(* IEC 61131-3 sources: TetherPLC/tests/compat, 95 files *)

(* ---- mqtt_blocks_case.st ---- *)
// mqtt_blocks_case.st — easy FBD blocks e2e: FB_MqttLink (wss://)
// + FB_MqttSub + FB_MqttTx + FB_MqttRx loopback through the fake
// broker's --ws --tls mode.  mask %QD0 bits (expect 0x1f):
//   b0 link Connected     b3 rx HasMsg fields match
//   b1 sub Done seen      b4 rx MsgCnt>=1
//   b2 tx Done seen
PROGRAM mqtt_blocks_case
VAR
    lk : FB_MqttLink;
    tx : FB_MqttTx;
    sub : FB_MqttSub;
    rx : FB_MqttRx;
    st : INT;
    mask AT %QD0 : UDINT;
    gotMsg : BOOL;
    gotCnt : BOOL;
END_VAR
    // link config — wss:// self-signed + credentials
    lk.Execute := TRUE;
    lk.Host := 'localhost';
    lk.Port := 11888;
    lk.User := 'wsuser';
    lk.Pass := 'wspass';
    lk.ClientId := 'blocks-e2e';
    lk.ConnectMs := 5000;
    lk.Transport := 4;            // wss
    lk.UseTls := TRUE;
    lk.TlsInsecure := TRUE;
    lk.BackoffMin := 500;
    lk.BackoffMax := 2000;
    // sub/tx are level-driven: Execute high only during their step
    sub.Hdl := lk.Hdl;
    sub.Filter := 'fbd/test/#';
    sub.Qos := 0;
    sub.Execute := (st = 1);
    tx.Hdl := lk.Hdl;
    tx.Topic := 'fbd/test/1';
    tx.Payload := 'PING';
    tx.Qos := 0;
    tx.Retained := FALSE;
    tx.Execute := (st = 2);

    lk();
    sub();
    tx();
    rx.Hdl := lk.Hdl;
    rx();

    IF st = 0 THEN
        mask := 0;
        IF lk.Connected THEN
            mask := mask + 1;
            st := 1;
        END_IF;
        IF st < 90 AND lk.Err THEN st := 90; END_IF;
    END_IF;
    IF st = 1 THEN
        IF sub.Done THEN
            mask := mask + 2;
            st := 2;
        END_IF;
        IF st < 90 AND lk.Err THEN st := 90; END_IF;
    END_IF;
    IF st = 2 THEN
        IF tx.Done THEN
            mask := mask + 4;
            st := 3;
        END_IF;
        IF st < 90 AND (lk.Err OR tx.Err) THEN st := 90; END_IF;
    END_IF;
    IF st >= 3 AND st < 90 THEN
        // rx fields persist — edge-guard so bits latch once
        IF rx.MsgCnt > 0 AND rx.Topic = 'fbd/test/1'
           AND rx.Payload = 'PING' AND NOT gotMsg THEN
            mask := mask + 8;
            gotMsg := TRUE;
        END_IF;
        IF rx.MsgCnt >= 1 AND NOT gotCnt THEN
            mask := mask + 16;
            gotCnt := TRUE;
        END_IF;
        IF mask >= 31 THEN
            st := 6;
        END_IF;
        IF st < 90 AND rx.Err THEN st := 90; END_IF;
    END_IF;
    IF st >= 90 THEN
        mask := 16#DEAD;
    END_IF;
END_PROGRAM

(* ---- mqtt_journal_case.st ---- *)
// mqtt_journal_case.st — ST-side event journal e2e: FB_MqttLink +
// FB_MqttSub + FB_MqttRx feed FB_MqttEventLog; the fake broker injects
// three messages on jrn/# after the subscription lands.
// mask %QD0 bits (expect 0x3f):
//   b0 link Connected     b3 LOG[0..2] topics+payloads in order
//   b1 sub Done seen      b4 journal Head entry = newest
//   b2 journal Count>=3   b5 rx MsgCnt>=3
PROGRAM mqtt_journal_case
VAR
    lk : FB_MqttLink;
    sub : FB_MqttSub;
    rx : FB_MqttRx;
    lg : FB_MqttEventLog;
    st : INT;
    mask AT %QD0 : UDINT;
    gotCnt : BOOL;
    gotRx : BOOL;
    gotTopics : BOOL;
    gotHead : BOOL;
    i : UDINT;
    nScan : UDINT;
    sawA : BOOL;
    sawB : BOOL;
    sawC : BOOL;
END_VAR
    lk.Execute := TRUE;
    lk.Host := 'localhost';
    lk.Port := 11883;
    lk.ClientId := 'journal-e2e';
    lk.ConnectMs := 5000;
    lk.BackoffMin := 500;
    lk.BackoffMax := 2000;

    sub.Hdl := lk.Hdl;
    sub.Filter := 'jrn/#';
    sub.Qos := 0;
    sub.Execute := (st = 1);

    rx.Hdl := lk.Hdl;
    lg.Execute := TRUE;
    lg.CycleTime := 0.01;
    lg.Push := rx.HasMsg;
    lg.TopicIn := rx.Topic;
    lg.PayloadIn := rx.Payload;

    lk();
    sub();
    rx();
    lg();

    IF st = 0 THEN
        mask := 0;
        IF lk.Connected THEN
            mask := mask + 1;
            st := 1;
        END_IF;
        IF st < 90 AND lk.Err THEN st := 90; END_IF;
    END_IF;
    IF st = 1 THEN
        IF sub.Done THEN
            mask := mask + 2;
            st := 2;
        END_IF;
        IF st < 90 AND lk.Err THEN st := 90; END_IF;
    END_IF;
    IF st >= 2 AND st < 90 THEN
        // journal content — injects repeat cyclically so arrival
        // order interleaves; require all three pairs present in the
        // ring (any order) rather than a fixed first-3 sequence
        IF lg.Count >= 3 AND NOT gotCnt THEN
            mask := mask + 4;
            gotCnt := TRUE;
        END_IF;
        IF lg.Count >= 3 AND NOT gotTopics THEN
            sawA := FALSE; sawB := FALSE; sawC := FALSE;
            nScan := lg.Count;
            IF nScan > 16 THEN nScan := 16; END_IF;
            FOR i := 0 TO 15 DO
                IF i < nScan THEN
                    IF lg.LOG[i].Topic = 'jrn/a'
                       AND lg.LOG[i].Payload = 'MSG1' THEN sawA := TRUE; END_IF;
                    IF lg.LOG[i].Topic = 'jrn/b'
                       AND lg.LOG[i].Payload = 'MSG2' THEN sawB := TRUE; END_IF;
                    IF lg.LOG[i].Topic = 'jrn/c'
                       AND lg.LOG[i].Payload = 'MSG3' THEN sawC := TRUE; END_IF;
                END_IF;
            END_FOR;
            IF sawA AND sawB AND sawC THEN
                mask := mask + 8;
                gotTopics := TRUE;
            END_IF;
        END_IF;
        IF lg.Count >= 1 AND NOT gotHead THEN
            // Head points at the newest entry — payload must be one
            // of the injected values and Tick must be > 0
            IF (lg.LOG[lg.Head].Payload = 'MSG1'
                OR lg.LOG[lg.Head].Payload = 'MSG2'
                OR lg.LOG[lg.Head].Payload = 'MSG3')
               AND lg.LOG[lg.Head].Tick > 0.0 THEN
                mask := mask + 16;
                gotHead := TRUE;
            END_IF;
        END_IF;
        IF rx.MsgCnt >= 3 AND NOT gotRx THEN
            mask := mask + 32;
            gotRx := TRUE;
        END_IF;
        // all bits latched → done (expect 0x3f)
        IF mask >= 63 THEN st := 90; END_IF;
    END_IF;
END_PROGRAM

(* ---- mqtt_tls_case.st ---- *)
// mqtt_tls_case.st — FB_Mqtt TLS e2e against the python fake broker
// (--tls).  Two sequential connects on one handle:
//   conn1: ssl:// + tls_insecure (self-signed accepted) + credentials
//   conn2: ssl:// + CA-file verification (TlsCaFile) + credentials
// mask %QD0 bits (expect 0x0f):
//   b0 conn1 CONNECTED    b2 conn2 CONNECTED
//   b1 conn1 publish ok   b3 conn2 publish ok
PROGRAM mqtt_tls_case
VAR
    m : FB_Mqtt;
    st : INT;
    mask AT %QD0 : UDINT;
    hdl : UDINT;
    caf : STRING[255];
END_VAR
    caf := '/tmp/tether_mqtt_tls/ca.pem';
    IF st = 0 THEN
        mask := 0;
        // ---- conn1: TLS, insecure (self-signed), creds, MQTT5 ----
        m.OP := 1;
        m.HOST := 'localhost';
        m.PORT := 11886;
        m.USERNAME := 'tlsuser';
        m.PASSWORD := 'tlspass';
        m.CLIENTID := 'tls-e2e-1';
        m.CONNECTMS := 3000;
        m.MQTTVER := 5;
        m.USETLS := 1;
        m.TLSINSECURE := 1;
        m.TLSCAFILE := '';
        m();
        IF m.STATUS = 0 THEN
            hdl := m.HANDLE;
            st := 1;
        ELSE
            st := 90;
        END_IF;
    END_IF;

    IF st = 1 THEN
        m.OP := 8;
        m.HANDLE := hdl;
        m();
        IF m.CONNECTED <> 0 THEN
            mask := mask + 1;
            st := 2;
        END_IF;
        IF st < 90 AND m.STATUS < 0 THEN st := 90; END_IF;
    END_IF;

    IF st = 2 THEN
        m.OP := 4;
        m.HANDLE := hdl;
        m.TOPIC := 'tls/one';
        m.PAYLOAD := 'A';
        m.QOS := 0;
        m.FLG_RETAIN := 0;
        m();
        IF m.STATUS = 0 THEN mask := mask + 2; END_IF;
        st := 3;
    END_IF;

    IF st = 3 THEN
        m.OP := 2;
        m.HANDLE := hdl;
        m();
        // ---- conn2: TLS with CA verification ----
        m.OP := 1;
        m.HOST := 'localhost';
        m.PORT := 11886;
        m.USERNAME := 'tlsuser';
        m.PASSWORD := 'tlspass';
        m.CLIENTID := 'tls-e2e-2';
        m.CONNECTMS := 3000;
        m.MQTTVER := 5;
        m.USETLS := 1;
        m.TLSINSECURE := 0;
        m.TLSCAFILE := caf;
        m();
        IF m.STATUS = 0 THEN
            hdl := m.HANDLE;
            st := 4;
        ELSE
            st := 90;
        END_IF;
    END_IF;

    IF st = 4 THEN
        m.OP := 8;
        m.HANDLE := hdl;
        m();
        IF m.CONNECTED <> 0 THEN
            mask := mask + 4;
            st := 5;
        END_IF;
        IF st < 90 AND m.STATUS < 0 THEN st := 90; END_IF;
    END_IF;

    IF st = 5 THEN
        m.OP := 4;
        m.HANDLE := hdl;
        m.TOPIC := 'tls/two';
        m.PAYLOAD := 'B';
        m.QOS := 0;
        m.FLG_RETAIN := 0;
        m();
        IF m.STATUS = 0 THEN mask := mask + 8; END_IF;
        st := 6;
    END_IF;

    IF st >= 90 THEN
        mask := 16#DEAD;
    END_IF;
END_PROGRAM

(* ---- mqtt_ws_case.st ---- *)
// mqtt_ws_case.st — FB_Mqtt WebSocket e2e against the python fake
// broker (--ws).  Two sequential connects:
//   conn1: ws://  (plain WebSocket, port 11887)
//   conn2: wss:// (WebSocket over TLS, self-signed, port 11888)
// Both carry username/password/client_id.  mask %QD0 bits
// (expect 0x0f):
//   b0 ws  CONNECTED    b2 wss CONNECTED
//   b1 ws  publish ok   b3 wss publish ok
PROGRAM mqtt_ws_case
VAR
    m : FB_Mqtt;
    st : INT;
    mask AT %QD0 : UDINT;
    hdl : UDINT;
    caf : STRING[255];
END_VAR
    caf := '/tmp/tether_mqtt_tls/ca.pem';
    IF st = 0 THEN
        mask := 0;
        // ---- conn1: ws:// plain WebSocket ----
        m.OP := 1;
        m.HOST := 'localhost';
        m.PORT := 11887;
        m.USERNAME := 'wsuser';
        m.PASSWORD := 'wspass';
        m.CLIENTID := 'ws-e2e-1';
        m.CONNECTMS := 5000;
        m.TRANSPORT := 3;             // ws
        m();
        IF m.STATUS = 0 THEN
            hdl := m.HANDLE;
            st := 1;
        ELSE
            st := 90;
        END_IF;
    END_IF;

    IF st = 1 THEN
        m.OP := 8;
        m.HANDLE := hdl;
        m();
        IF m.CONNECTED <> 0 THEN
            mask := mask + 1;
            st := 2;
        END_IF;
        IF st < 90 AND m.STATUS < 0 THEN st := 90; END_IF;
    END_IF;

    IF st = 2 THEN
        m.OP := 4;
        m.HANDLE := hdl;
        m.TOPIC := 'ws/one';
        m.PAYLOAD := 'A';
        m.QOS := 0;
        m.FLG_RETAIN := 0;
        m();
        IF m.STATUS = 0 THEN mask := mask + 2; END_IF;
        st := 3;
    END_IF;

    IF st = 3 THEN
        m.OP := 2;
        m.HANDLE := hdl;
        m();
        // ---- conn2: wss:// WebSocket over TLS (self-signed) ----
        m.OP := 1;
        m.HOST := 'localhost';
        m.PORT := 11888;
        m.USERNAME := 'wsuser';
        m.PASSWORD := 'wspass';
        m.CLIENTID := 'ws-e2e-2';
        m.CONNECTMS := 5000;
        m.TRANSPORT := 4;             // wss
        m.USETLS := 1;
        m.TLSINSECURE := 1;
        m.TLSCAFILE := '';
        m();
        IF m.STATUS = 0 THEN
            hdl := m.HANDLE;
            st := 4;
        ELSE
            st := 90;
        END_IF;
    END_IF;

    IF st = 4 THEN
        m.OP := 8;
        m.HANDLE := hdl;
        m();
        IF m.CONNECTED <> 0 THEN
            mask := mask + 4;
            st := 5;
        END_IF;
        IF st < 90 AND m.STATUS < 0 THEN st := 90; END_IF;
    END_IF;

    IF st = 5 THEN
        m.OP := 4;
        m.HANDLE := hdl;
        m.TOPIC := 'ws/two';
        m.PAYLOAD := 'B';
        m.QOS := 0;
        m.FLG_RETAIN := 0;
        m();
        IF m.STATUS = 0 THEN mask := mask + 8; END_IF;
        st := 6;
    END_IF;

    IF st >= 90 THEN
        mask := 16#DEAD;
    END_IF;
END_PROGRAM

(* ---- tc2_aes70_case.st ---- *)
// tc2_aes70_case.st — OCA/AES70 client e2e over the python device
// fake.  Connect, keepalive, a method call -> echoed response,
// disconnect.
PROGRAM tc2_aes70_case
VAR
    con : FB_Aes70Connect;
    dis : FB_Aes70Disconnect;
    ka  : FB_Aes70Keepalive;
    cal : FB_Aes70Call;
    rx  : FB_Aes70Receive;
    st : INT;
    waitN : INT;
    mask AT %QD0 : UDINT;
    hdl : UDINT;
END_VAR
    IF st = 0 THEN
        mask := 0;
        con.Execute := TRUE;
        con.Host := '127.0.0.1';
        con.Port := 65000;
        st := 1;
    END_IF;

    IF st = 1 THEN
        IF con.Done THEN
            hdl := con.ConnectionHdl;
            con.Execute := FALSE;
            mask := mask + 1;         // bit0: session up
            ka.Execute := TRUE;
            ka.ConnectionHdl := hdl;
            st := 2;
        END_IF;
        IF con.Error THEN mask := 16#DEAD; st := 99; END_IF;
    END_IF;

    IF st = 2 THEN
        IF ka.Done THEN
            mask := mask + 2;         // bit1: keepalive sent
            ka.Execute := FALSE;
            cal.Execute := TRUE;
            cal.ConnectionHdl := hdl;
            cal.TargetONo := 1000;    // an OCA object number
            cal.MethodID := 260;      // defLevel=1, methodIndex=4
            cal.Params := '{"gain":0.5}';
            st := 3;
        END_IF;
        IF ka.Error THEN mask := 16#DEAD; st := 99; END_IF;
    END_IF;

    IF st = 3 THEN
        IF cal.Done THEN
            mask := mask + 4;         // bit2: call sent
            cal.Execute := FALSE;
            rx.Execute := TRUE;
            rx.ConnectionHdl := hdl;
            st := 4;
        END_IF;
        IF cal.Error THEN mask := 16#DEAD; st := 99; END_IF;
    END_IF;

    // poll for the device's echoed OcaResponse
    IF st = 4 THEN
        waitN := waitN + 1;
        IF rx.Message THEN
            mask := mask + 8;         // bit3: response landed
            rx.Execute := FALSE;
            dis.Execute := TRUE;
            dis.ConnectionHdl := hdl;
            st := 5;
        END_IF;
        IF rx.Error THEN mask := 16#DEAD; st := 99; END_IF;
        IF waitN > 40 THEN
            rx.Execute := FALSE;
            dis.Execute := TRUE;
            dis.ConnectionHdl := hdl;
            st := 5;
        END_IF;
    END_IF;

    IF st = 5 THEN
        IF dis.Done THEN
            mask := mask + 16;        // bit4: released
            st := 6;
        END_IF;
        IF dis.Error THEN mask := 16#DEAD; st := 99; END_IF;
    END_IF;

    con(); dis(); ka(); cal(); rx();
END_PROGRAM

(* ---- tc2_babasic_case.st ---- *)
// tc2_babasic_case.st — pure-ST e2e for tc2_babasic.
// Exercises the core blocks; mask bits land per check.
PROGRAM tc2_babasic_case
VAR
    thr : FB_ThresholdSwitch;
    ramp : FB_Ramp;
    lgt : FB_Light;
    stair : FB_StairwellLight;
    mdc : FB_MaximumDemandController;
    sched : FB_DailyScheduler;
    scn : FB_ScenesLighting;
    scl : LREAL;
    st : INT;
    mask AT %QD0 : UDINT;
    diag AT %QD4 : UDINT;
END_VAR
    diag := st;
    IF st = 0 THEN
        mask := 0;
        // F_Scale: 50 in 0..100 -> 0..10 = 5
        scl := F_Scale(50.0, 0.0, 100.0, 0.0, 10.0);
        IF scl > 4.9 AND scl < 5.1 THEN mask := mask OR 1; END_IF;
        st := 1;
    ELSIF st = 1 THEN
        thr.x := 10.0; thr.On := 5.0; thr.Off := 1.0;
        thr();
        IF thr.Q THEN mask := mask OR 2; END_IF;
        st := 2;
    ELSIF st = 2 THEN
        ramp.Enable := TRUE;
        ramp.Setpoint := 10.0;
        ramp.SlewUp := 5.0;
        ramp.SlewDown := 5.0;
        ramp.CycleTime := 0.1;
        IF ramp.Out > 0.4 THEN mask := mask OR 4; st := 3; END_IF;
    ELSIF st = 3 THEN
        // run ramp to target over 25 scans
        diag := diag + 0;         // keep diag = st
        IF ramp.AtTarget THEN mask := mask OR 8; st := 4; END_IF;
    ELSIF st = 4 THEN
        lgt.On := TRUE;
        lgt.OffDelay := 0.3;
        lgt.CycleTime := 0.1;
        IF lgt.Q THEN mask := mask OR 16; st := 5; END_IF;
    ELSIF st = 5 THEN
        stair.Trigger := TRUE;
        stair.Duration := 0.5;
        stair.CycleTime := 0.1;
        IF stair.Q THEN mask := mask OR 32; st := 6; END_IF;
    ELSIF st = 6 THEN
        mdc.Enable := TRUE;
        mdc.In1 := TRUE; mdc.In2 := TRUE; mdc.In3 := TRUE; mdc.In4 := TRUE;
        mdc.Limit := 2;
        st := 7;
    ELSIF st = 7 THEN
        IF mdc.Shedding AND mdc.Q1 AND mdc.Q2 AND NOT mdc.Q3 AND NOT mdc.Q4 THEN
            mask := mask OR 64;
        END_IF;
        sched.Enable := TRUE;
        sched.MinuteOfDay := 700;   // 11:40
        sched.OnMin := 600;         // 10:00
        sched.OffMin := 720;        // 12:00
        scn.Enable := TRUE;
        scn.Scene := 2;
        scn.L2 := 77.0;
        st := 8;
    ELSIF st = 8 THEN
        IF sched.Q AND scn.Q AND scn.Level = 77.0 THEN
            mask := mask OR 128;
        END_IF;
        st := 9;
    END_IF;
    thr(); ramp(); lgt(); stair(); mdc(); sched(); scn();
END_PROGRAM

(* ---- tc2_case.st ---- *)
PROGRAM Tc2Case
VAR
    start_in AT %IX0.0 : BOOL;
    mask      AT %QD0   : DINT;
    tmask     AT %QD4   : DINT;
    d2b       : DEC_TO_BCD;
    b2d       : BCD_TO_DEC;
    d2b_err   : DEC_TO_BCD;
    lton1     : LTON;
    ltof1     : LTOF;
    ltp1      : LTP;
    enm       : FB_EnumStringNumbers;
    enm2      : FB_EnumStringNumbers;
    enm3      : FB_EnumStringNumbers;
    scan_n    : UDINT;
    eCmd      : INT;
END_VAR

d2b(START := start_in, DIN := 42);
b2d(START := start_in, BIN := 16#26);
d2b_err(START := start_in, DIN := 200);
lton1(IN := start_in, PT := T#15ms);
ltof1(IN := start_in, PT := T#20ms);
ltp1(IN := start_in, PT := T#25ms);
IF scan_n = 0 THEN
    eCmd := 0;
ELSE
    eCmd := 1;
END_IF
enm(sSearch := 'abc12.5xyz-7', eCmd := eCmd, eType := 0);
enm2(sSearch := 'abc12.5xyz', eCmd := 0, eType := 0);
enm3(sSearch := '-7x', eCmd := 0, eType := 2);
scan_n := scan_n + 1;

mask := 0;
IF CEIL(2.3) = 3.0 THEN
    mask := mask + 1;
END_IF
IF FLOOR(-2.3) = -3.0 THEN
    mask := mask + 2;
END_IF
IF FRAC(3.25) = 0.25 THEN
    mask := mask + 4;
END_IF
IF LTRUNC(-3.7) = -3.0 THEN
    mask := mask + 8;
END_IF
IF LMOD(7.5, 2.0) = 1.5 THEN
    mask := mask + 16;
END_IF
IF MODABS(-7.5, 2.0) = 0.5 THEN
    mask := mask + 32;
END_IF
IF MODTURNS(7.5, 2.0) = 3 THEN
    mask := mask + 64;
END_IF
IF MODTURNS(-7.5, 2.0) = -3 THEN
    mask := mask + 128;
END_IF
IF WCONCAT("ab", "cd") = "abcd" THEN
    mask := mask + 256;
END_IF
IF WLEFT("hello", 2) = "he" THEN
    mask := mask + 512;
END_IF
IF WRIGHT("hello", 2) = "lo" THEN
    mask := mask + 1024;
END_IF
IF WMID("hello", 3, 2) = "ell" THEN
    mask := mask + 2048;
END_IF
IF WFIND("hello", "ll") = 3 THEN
    mask := mask + 4096;
END_IF
IF WLEN("hello") = 5 THEN
    mask := mask + 8192;
END_IF
IF WINSERT("ac", "b", 2) = "abc" THEN
    mask := mask + 16384;
END_IF
IF WDELETE("abc", 1, 2) = "ac" THEN
    mask := mask + 32768;
END_IF
IF WREPLACE("abc", "x", 1, 2) = "axc" THEN
    mask := mask + 65536;
END_IF
IF d2b.BOUT = 16#42 THEN
    mask := mask + 131072;
END_IF
IF b2d.DOUT = 26 THEN
    mask := mask + 262144;
END_IF
IF d2b_err.ERR THEN
    mask := mask + 524288;
END_IF
IF d2b_err.ERRID <> 0 THEN
    mask := mask + 1048576;
END_IF

tmask := 0;
IF lton1.Q = FALSE THEN
    tmask := tmask + 1;
END_IF
IF ltof1.Q = TRUE THEN
    tmask := tmask + 2;
END_IF
IF ltp1.Q = FALSE THEN
    tmask := tmask + 4;
END_IF
IF enm2.sNumber = '12.5' THEN
    tmask := tmask + 8;
END_IF
IF enm3.sNumber = '-7' THEN
    tmask := tmask + 16;
END_IF
IF enm.bEOS = TRUE THEN
    tmask := tmask + 32;
END_IF
IF enm.nPos = 13 THEN
    tmask := tmask + 64;
END_IF
IF enm2.nPos = 8 THEN
    tmask := tmask + 128;
END_IF
END_PROGRAM

(* ---- tc2_cm_case.st ---- *)
// tc2_cm_case.st — CM e2e: function generator, linear interp,
// cam profile — pure-ST curve/math.
PROGRAM tc2_cm_case
VAR
    fg : FB_FuncGen;
    li : FB_LinInterp;
    cam : FB_CamProfile;
    st : INT;
    n : INT;
    mask AT %QD0 : UDINT;
END_VAR
    IF st = 0 THEN
        mask := 0;
        fg.Execute := TRUE;
        li.Execute := TRUE;
        cam.Execute := TRUE;
        fg.Shape := 1;            // triangle
        fg.Period := 1.0;
        fg.Amplitude := 2.0;
        fg.Offset := 0.0;
        fg.CycleTime := 0.1;
        li.X := 1.5;
        li.X0 := 0.0; li.Y0 := 0.0;
        li.X1 := 1.0; li.Y1 := 2.0;
        li.X2 := 2.0; li.Y2 := 4.0;
        li.X3 := 3.0; li.Y3 := 8.0;
        cam.MasterEnd := 10.0;
        cam.SlaveAmp := 100.0;
        cam.Master := 5.0;
        st := 1;
    END_IF;

    // funcgen runs — phase advances
    IF st = 1 THEN
        IF fg.Done THEN
            n := n + 1;
            IF n > 8 THEN
                IF fg.Phase > 0.0 THEN mask := mask + 1; END_IF;
                n := 0;
                st := 2;
            END_IF;
        END_IF;
    END_IF;
    // lininterp X=1.5 between (1,2)->(2,4) -> Y=3
    IF st = 2 THEN
        IF li.Done THEN
            IF li.Y > 2.9 AND li.Y < 3.1 THEN mask := mask + 2; END_IF;
            st := 3;
        END_IF;
    END_IF;
    // cam: master 5 of 10 -> slave ~50 of 100
    IF st = 3 THEN
        IF cam.Done THEN
            IF cam.Slave > 49.0 AND cam.Slave < 51.0 THEN
                mask := mask + 4;
            END_IF;
            IF cam.InSync THEN mask := mask + 8; END_IF;
            st := 4;
        END_IF;
    END_IF;
    // funcgen output in range
    IF st = 4 THEN
        IF fg.Done THEN
            IF fg.Output >= 0.0 AND fg.Output <= 2.0 THEN
                mask := mask + 16;
            END_IF;
            st := 5;
        END_IF;
    END_IF;

    fg(); li(); cam();
END_PROGRAM

(* ---- tc2_ctb_case.st ---- *)
// tc2_ctb_case.st — Tc2_ControllerToolbox e2e: hysteresis, two-
// position, deadtime, statistics, PWM — pure-ST blocks.
PROGRAM tc2_ctb_case
VAR
    hys : FB_Hysteresis;
    two : FB_TwoPosition;
    dt  : FB_DeadTime;
    stt : FB_Statistics;
    pwm : FB_Pwm;
    st : INT;
    n : INT;
    mask AT %QD0 : UDINT;
END_VAR
    IF st = 0 THEN
        mask := 0;
        hys.Execute := TRUE;
        two.Execute := TRUE;
        dt.Execute := TRUE;
        stt.Execute := TRUE;
        pwm.Execute := TRUE;
        hys.Input := 0.5; hys.OnLevel := 0.3; hys.OffLevel := 0.8;
        two.Setpoint := 1.0; two.Actual := 0.0; two.Hysteresis := 0.2;
        dt.Input := 7.0; dt.DelayCycles := 3;
        stt.Input := 2.0; stt.N := 4;
        pwm.Duty := 50.0; pwm.Period := 1.0; pwm.CycleTime := 0.1;
        st := 1;
    END_IF;

    // hysteresis: 0.5 is between 0.3..0.8 — stays off (started off)
    IF st = 1 THEN
        IF hys.Done THEN
            IF hys.Out = FALSE THEN mask := mask + 1; END_IF;
            st := 2;
        END_IF;
    END_IF;
    // two-position: Actual 0 < SP 1 - hyst -> drive on
    IF st = 2 THEN
        IF two.Done THEN
            IF two.Out = TRUE THEN mask := mask + 2; END_IF;
            st := 3;
        END_IF;
    END_IF;
    // deadtime: after DelayCycles the output lags input
    IF st = 3 THEN
        IF dt.Done THEN
            n := n + 1;
            IF n > 6 THEN
                IF dt.Output = 7.0 THEN mask := mask + 4; END_IF;
                n := 0;
                st := 4;
            END_IF;
        END_IF;
    END_IF;
    // statistics: mean of constant input ~= input, stddev ~0
    IF st = 4 THEN
        IF stt.Done THEN
            n := n + 1;
            IF n > 8 THEN
                IF stt.Mean > 1.9 AND stt.StdDev < 0.2 THEN
                    mask := mask + 8;
                END_IF;
                n := 0;
                st := 5;
            END_IF;
        END_IF;
    END_IF;
    // pwm: 50% duty -> Out toggles; just verify it ran
    IF st = 5 THEN
        IF pwm.Done THEN
            mask := mask + 16;
            st := 6;
        END_IF;
    END_IF;

    hys(); two(); dt(); stt(); pwm();
END_PROGRAM

(* ---- tc2_dataexchange_case.st ---- *)
// tc2_dataexchange_case.st — e2e for tc2_dataexchange (tplc-sym).
// The program's own variables are addressed by name through the
// package's exported var table.
PROGRAM tc2_dataexchange_case
VAR
    rd : FB_ReadAdsSymByName;
    wr : FB_WriteAdsSymByName;
    dI : FB_WriteDWordOnDelta;
    dR : FB_WriteLRealOnDelta;
    wd : FB_CheckWatchdog;
    heartbeat : DINT;
    setpoint : LREAL;
    flag : BOOL;
    st : INT;
    mask AT %QD0 : UDINT;
    diag AT %QD4 : UDINT;
END_VAR
    diag := st;
    IF st = 0 THEN
        mask := 0;
        wr.sVarName := 'heartbeat';
        wr.nIntValue := 1234;
        wr.bWrite := TRUE;
        st := 1;
    ELSIF st = 1 THEN
        IF wr.bDone THEN mask := mask OR 1; END_IF;
        wr.bWrite := FALSE;
        IF heartbeat = 1234 THEN mask := mask OR 2; END_IF;
        rd.sVarName := 'heartbeat';
        st := 2;
    ELSIF st = 2 THEN
        rd.bRead := TRUE;
        st := 3;
    ELSIF st = 3 THEN
        IF rd.nIntValue = 1234 AND rd.nSize = 4 THEN mask := mask OR 4; END_IF;
        rd.bRead := FALSE;
        wr.sVarName := 'setpoint';
        wr.fRealValue := 12.5;
        st := 4;
    ELSIF st = 4 THEN
        wr.bWrite := TRUE;
        st := 5;
    ELSIF st = 5 THEN
        IF wr.bDone AND setpoint = 12.5 THEN mask := mask OR 8; END_IF;
        wr.bWrite := FALSE;
        wr.sVarName := 'flag';
        wr.bBoolValue := TRUE;
        st := 6;
    ELSIF st = 6 THEN
        wr.bWrite := TRUE;
        st := 7;
    ELSIF st = 7 THEN
        IF wr.bDone AND flag THEN mask := mask OR 16; END_IF;
        wr.bWrite := FALSE;
        // unknown name must error
        wr.sVarName := 'no_such_var';
        st := 8;
    ELSIF st = 8 THEN
        wr.bWrite := TRUE;
        st := 9;
    ELSIF st = 9 THEN
        IF wr.bError THEN mask := mask OR 32; END_IF;
        wr.bWrite := FALSE;
        // delta writer: transmits on change only
        dI.sVarName := 'heartbeat';
        dI.nValue := 7;
        st := 10;
    ELSIF st = 10 THEN
        dI.bEnable := TRUE;
        st := 11;
    ELSIF st = 11 THEN
        IF dI.nLastSignal = 7 AND heartbeat = 7 THEN mask := mask OR 64; END_IF;
        dR.sVarName := 'setpoint';
        dR.fValue := 3.25;
        st := 12;
    ELSIF st = 12 THEN
        dR.bEnable := TRUE;
        st := 13;
    ELSIF st = 13 THEN
        IF dR.fLastSignal = 3.25 AND setpoint = 3.25 THEN
            mask := mask OR 128;
        END_IF;
        // watchdog: heartbeat is written every scan by the delta
        // block?  No — use a dedicated stamp variable.
        wd.sVarName := 'heartbeat';
        wd.tTimeout := T#1S;
        st := 14;
    ELSIF st = 14 THEN
        wd.bEnable := TRUE;
        st := 15;
    ELSIF st = 15 THEN
        IF wd.bAlive AND NOT wd.bTimeout THEN mask := mask OR 256; END_IF;
        st := 16;
    END_IF;
    rd(); wr(); dI(); dR(); wd();
END_PROGRAM

(* ---- tc2_dmx_case.st ---- *)
// tc2_dmx_case.st — DMX512 output e2e over a PTY fake.  Open,
// set channels, send a frame, status, close.
PROGRAM tc2_dmx_case
VAR
    opn : FB_DmxOpen;
    cls : FB_DmxClose;
    set : FB_DmxSetChannel;
    snd : FB_DmxSend;
    sta : FB_DmxStatus;
    st : INT;
    waitN : INT;
    mask AT %QD0 : UDINT;
    hdl : UDINT;
END_VAR
    IF st = 0 THEN
        mask := 0;
        opn.Execute := TRUE;
        opn.Path := '/tmp/dmx_pty';
        opn.Baud := 250000;
        st := 1;
    END_IF;

    IF st = 1 THEN
        IF opn.Done THEN
            hdl := opn.PortHdl;
            opn.Execute := FALSE;
            mask := mask + 1;         // bit0: serial open
            set.Execute := TRUE;
            set.PortHdl := hdl;
            set.Channel := 1;
            set.Value := 200;
            st := 2;
        END_IF;
        IF opn.Error THEN mask := 16#DEAD; st := 99; END_IF;
    END_IF;

    IF st = 2 THEN
        IF set.Done THEN
            mask := mask + 2;         // bit1: channel written
            set.Execute := FALSE;
            snd.Execute := TRUE;
            snd.PortHdl := hdl;
            st := 3;
        END_IF;
        IF set.Error THEN mask := 16#DEAD; st := 99; END_IF;
    END_IF;

    IF st = 3 THEN
        IF snd.Done THEN
            mask := mask + 4;         // bit2: frame emitted
            snd.Execute := FALSE;
            sta.Execute := TRUE;
            sta.PortHdl := hdl;
            st := 4;
        END_IF;
        IF snd.Error THEN mask := 16#DEAD; st := 99; END_IF;
    END_IF;

    IF st = 4 THEN
        IF sta.Done THEN
            IF sta.Frames > 0 THEN
                mask := mask + 8;     // bit3: frame counted
            END_IF;
            sta.Execute := FALSE;
            cls.Execute := TRUE;
            cls.PortHdl := hdl;
            st := 5;
        END_IF;
        IF sta.Error THEN mask := 16#DEAD; st := 99; END_IF;
    END_IF;

    IF st = 5 THEN
        IF cls.Done THEN
            mask := mask + 16;        // bit4: closed
            st := 6;
        END_IF;
        IF cls.Error THEN mask := 16#DEAD; st := 99; END_IF;
    END_IF;

    opn(); cls(); set(); snd(); sta();
END_PROGRAM

(* ---- tc2_drive_case.st ---- *)
// tc2_drive_case.st — Tc2_Drive e2e over the Tether IO backend.
// Exercises the SoE surface (state read, diag fields, password,
// command control/exec/state, error+reset, AX5000 blocks) against
// tether_io_motion_server's ec.soe.* params, plus the
// SimplePlcMotion CoE/SoE enable + velocity blocks on a simulated
// CiA402 axis. 14 checks packed into %QD0; last step expects
// mask 0x3fff.
PROGRAM tc2_drive_case
VAR
    mask   AT %QD0 : DINT;
    st     : INT;
    ph     : INT;
    wrN    : INT;
    cur    : INT;
    tgl    : BOOL;
    axH    : UDINT;
    pos    : DINT;

    ax     : FB_MotionAxis;
    axC    : FB_MotionAxis;

    stFb   : FB_SoEReadStatus;
    msgFb  : FB_SoEReadDiagMessage;
    numFb  : FB_SoEReadDiagNumber;
    lstFb  : FB_SoEReadDiagNumberList;
    clsFb  : FB_SoEReadClassXDiag;
    atFb   : FB_SoEReadAmplifierTemperature;
    mtFb   : FB_SoEReadMotorTemperature;
    dvFb   : FB_SoEReadDcBusVoltage;
    dcFb   : FB_SoEReadDcBusCurrent;
    pwFb   : FB_SoEWritePassword;
    ccFb   : FB_SoEWriteCommandControl;
    exFb   : FB_SoEExecuteCommand;
    rsFb   : FB_SoEReset;
    vmFb   : FB_SoEAX5000ReadActMainVoltage;
    mcFb   : FB_SoEAX5000SetMotorCtrlWord;
    fwFb   : FB_SoEAX5000FirmwareUpdate;
    pkFb   : FB_SoEAX5000ParkAxis;
    enFb   : FB_CoEDriveEnable;
    mvFb   : FB_SoEDriveMoveVelocity;
END_VAR

cur := st;

// ---- st=0: create the motion axis (for SimplePlcMotion) ----
IF cur = 0 THEN
    mask := 0;
    ph := 0;
    wrN := 0;
    tgl := FALSE;
    ax.UNITS_PER_REV := 1000;
    ax.MAX_VEL := 4000;
    ax.MAX_ACCEL := 20000;
    ax.MAX_DECEL := 20000;
    ax.POS_MIN := -100000;
    ax.POS_MAX := 100000;
    ax.HOME_OFFSET := 0;
    ax.FOLLOW_WINDOW := 10;
    ax.FLAGS := 1;
    ax.OP := 1; ax();
    axH := ax.AXIS;
    st := 1;
END_IF;

// ---- st=1: axis created? ----
IF cur = 1 THEN
    IF axH <> 0 THEN
        mask := mask + 1;          // bit0
        st := 2;
    ELSIF wrN > 50 THEN
        st := 90;
    ELSE
        wrN := wrN + 1;
    END_IF;
END_IF;

// ---- st=2/3: SoE status read (slave 0) ----
IF cur = 2 THEN
    stFb.Drive := 0;
    stFb.Execute := TRUE;
    st := 3;
END_IF;
IF cur = 3 THEN
    stFb.Execute := FALSE;
    IF stFb.bDone AND stFb.StatusWord = 3 AND stFb.CommandState = 0 THEN
        mask := mask + 2;          // bit1
    END_IF;
    st := 4;
END_IF;

// ---- st=4/5: diag number + list + class-X (slave 0) ----
IF cur = 4 THEN
    numFb.Drive := 0; numFb.Execute := TRUE;
    lstFb.Drive := 0; lstFb.Execute := TRUE;
    clsFb.Drive := 0; clsFb.Execute := TRUE;
    st := 5;
END_IF;
IF cur = 5 THEN
    numFb.Execute := FALSE;
    lstFb.Execute := FALSE;
    clsFb.Execute := FALSE;
    IF numFb.bDone AND numFb.DiagNumber = 16#8105 AND
       clsFb.bDone AND clsFb.ClassXDiag = 3 AND
       lstFb.bDone AND lstFb.DiagCount = 3 AND
       lstFb.DiagList[0] = 16#8105 THEN
        mask := mask + 4;          // bit2
    END_IF;
    st := 6;
END_IF;

// ---- st=6/7: diag message + temperatures + bus values ----
IF cur = 6 THEN
    msgFb.Drive := 0; msgFb.Execute := TRUE;
    atFb.Drive := 0;  atFb.Execute := TRUE;
    mtFb.Drive := 0;  mtFb.Execute := TRUE;
    dvFb.Drive := 0;  dvFb.Execute := TRUE;
    dcFb.Drive := 0;  dcFb.Execute := TRUE;
    st := 7;
END_IF;
IF cur = 7 THEN
    msgFb.Execute := FALSE;
    atFb.Execute := FALSE;
    mtFb.Execute := FALSE;
    dvFb.Execute := FALSE;
    dcFb.Execute := FALSE;
    IF msgFb.bDone AND msgFb.DiagMessage = 'OVERLOAD' AND
       atFb.bDone AND atFb.Value = 61.5 AND
       mtFb.bDone AND mtFb.Value = 58.25 AND
       dvFb.bDone AND dvFb.Value = 565.5 AND
       dcFb.bDone AND dcFb.Value = 12.75 THEN
        mask := mask + 8;          // bit3
    END_IF;
    st := 8;
END_IF;

// ---- st=8/9/10/11: password write, command-control write,
//      then one status re-read verifying both readbacks ----
IF cur = 8 THEN
    pwFb.Drive := 0;
    pwFb.Password := 16#1234;
    pwFb.Execute := TRUE;
    st := 9;
END_IF;
IF cur = 9 THEN
    pwFb.Execute := FALSE;
    ccFb.Drive := 0;
    ccFb.CommandControl := 16#55AA;
    ccFb.Execute := TRUE;
    st := 10;
END_IF;
IF cur = 10 THEN
    ccFb.Execute := FALSE;
    stFb.Drive := 0;
    stFb.Execute := TRUE;
    st := 11;
END_IF;
IF cur = 11 THEN
    stFb.Execute := FALSE;
    IF stFb.bDone AND stFb.Password = 16#1234 THEN
        mask := mask + 16;         // bit4
    END_IF;
    IF stFb.bDone AND stFb.CmdCtrl = 16#55AA THEN
        mask := mask + 32;         // bit5
    END_IF;
    st := 12;
END_IF;

// ---- st=12/13/14: execute command 0x0007, poll for done (2) ----
IF cur = 12 THEN
    exFb.Drive := 0;
    exFb.CommandId := 16#0007;
    exFb.Execute := TRUE;
    st := 13;
END_IF;
IF cur = 13 THEN
    exFb.Execute := FALSE;
    tgl := FALSE;
    wrN := 0;
    st := 14;
END_IF;
IF cur = 14 THEN
    tgl := NOT tgl;
    stFb.Drive := 0;
    stFb.Execute := tgl;
    IF stFb.bDone AND stFb.CommandState = 2 THEN
        mask := mask + 64;         // bit6
        stFb.Execute := FALSE;
        st := 15;
    ELSIF wrN > 80 THEN
        stFb.Execute := FALSE;
        st := 90;
    ELSE
        wrN := wrN + 1;
    END_IF;
END_IF;

// ---- st=15/16/17: execute command 0x8001 -> error state + fault ----
IF cur = 15 THEN
    exFb.Drive := 0;
    exFb.CommandId := 16#8001;
    exFb.Execute := TRUE;
    st := 16;
END_IF;
IF cur = 16 THEN
    exFb.Execute := FALSE;
    tgl := FALSE;
    wrN := 0;
    st := 17;
END_IF;
IF cur = 17 THEN
    tgl := NOT tgl;
    stFb.Drive := 0;
    stFb.Execute := tgl;
    IF stFb.bDone AND stFb.CommandState = 3 AND
       (stFb.StatusWord AND 4) <> 0 THEN
        mask := mask + 128;        // bit7
        stFb.Execute := FALSE;
        st := 18;
    ELSIF wrN > 80 THEN
        stFb.Execute := FALSE;
        st := 90;
    ELSE
        wrN := wrN + 1;
    END_IF;
END_IF;

// ---- st=18/19/20: reset clears the fault + command state ----
IF cur = 18 THEN
    rsFb.Drive := 0;
    rsFb.Execute := TRUE;
    st := 19;
END_IF;
IF cur = 19 THEN
    rsFb.Execute := FALSE;
    tgl := FALSE;
    wrN := 0;
    st := 20;
END_IF;
IF cur = 20 THEN
    tgl := NOT tgl;
    stFb.Drive := 0;
    stFb.Execute := tgl;
    IF stFb.bDone AND stFb.CommandState = 0 AND
       (stFb.StatusWord AND 4) = 0 THEN
        mask := mask + 256;        // bit8
        stFb.Execute := FALSE;
        st := 21;
    ELSIF wrN > 80 THEN
        stFb.Execute := FALSE;
        st := 90;
    ELSE
        wrN := wrN + 1;
    END_IF;
END_IF;

// ---- st=21..24: AX5000 motor ctrl word, park, mains, fw ----
IF cur = 21 THEN
    mcFb.Drive := 0;
    mcFb.MotorCtrlWord := 16#A5A5;
    mcFb.Execute := TRUE;
    st := 22;
END_IF;
IF cur = 22 THEN
    mcFb.Execute := FALSE;
    pkFb.Drive := 0;
    pkFb.Park := TRUE;
    pkFb.Execute := TRUE;
    st := 23;
END_IF;
IF cur = 23 THEN
    pkFb.Execute := FALSE;
    vmFb.Drive := 0; vmFb.Execute := TRUE;
    fwFb.Drive := 0; fwFb.Execute := TRUE;
    stFb.Drive := 0; stFb.Execute := TRUE;
    st := 24;
END_IF;
IF cur = 24 THEN
    vmFb.Execute := FALSE;
    fwFb.Execute := FALSE;
    stFb.Execute := FALSE;
    IF stFb.bDone AND stFb.AxCtrl = 16#A5A5 AND
       stFb.AxPark = 1 AND stFb.AxFwRev = 1 AND stFb.AxFwBuild = 5 AND
       vmFb.bDone AND vmFb.Voltage >= 230.0 AND vmFb.Voltage < 240.0 AND
       fwFb.bDone AND fwFb.FirmwareRevision = 1 AND
       fwFb.FirmwareBuild = 5 THEN
        mask := mask + 512;        // bit9
    END_IF;
    st := 25;
END_IF;

// ---- st=25/26: slave 1 diag number (OVERTEMP) ----
IF cur = 25 THEN
    numFb.Drive := 1;
    numFb.Execute := TRUE;
    st := 26;
END_IF;
IF cur = 26 THEN
    numFb.Execute := FALSE;
    IF numFb.bDone AND numFb.DiagNumber = 16#8201 THEN
        mask := mask + 1024;       // bit10
    END_IF;
    st := 27;
END_IF;

// ---- st=27/28: slave 5 has no diag entries ----
IF cur = 27 THEN
    lstFb.Drive := 5;
    lstFb.Execute := TRUE;
    st := 28;
END_IF;
IF cur = 28 THEN
    lstFb.Execute := FALSE;
    IF lstFb.bDone AND lstFb.DiagCount = 0 THEN
        mask := mask + 2048;       // bit11
    END_IF;
    st := 29;
END_IF;

// ---- st=29/30: CoE drive enable on the motion axis ----
IF cur = 29 THEN
    enFb.Enable := TRUE;
    enFb.Drive := axH;
    enFb.Execute := TRUE;
    st := 30;
END_IF;
IF cur = 30 THEN
    enFb.Execute := FALSE;
    IF enFb.bDone THEN
        mask := mask + 4096;       // bit12
    END_IF;
    mvFb.Drive := axH;
    mvFb.Velocity := 500.0;
    mvFb.Execute := TRUE;
    wrN := 0;
    st := 31;
END_IF;

// ---- st=31: SoE velocity move; wait for position > 50 ----
IF cur = 31 THEN
    axC.AXIS := axH;
    axC.OP := 4; axC.INDEX := 16#6064; axC();
    pos := axC.VALUE;
    IF pos > 50 THEN
        mask := mask + 8192;       // bit13
        mvFb.Execute := FALSE;
        st := 90;
    ELSIF wrN > 300 THEN
        mvFb.Execute := FALSE;
        st := 90;
    ELSE
        wrN := wrN + 1;
    END_IF;
END_IF;

// FB invocations (one call per scan each)
ax(); axC();
stFb(); msgFb(); numFb(); lstFb(); clsFb();
atFb(); mtFb(); dvFb(); dcFb();
pwFb(); ccFb(); exFb(); rsFb();
vmFb(); mcFb(); fwFb(); pkFb();
enFb(); mvFb();
END_PROGRAM

(* ---- tc2_eip_case.st ---- *)
// tc2_eip_case.st — EtherNet/IP client e2e over the fake adapter.
// ListIdentity, RegisterSession, Get/Set_Attribute_Single, close.
PROGRAM tc2_eip_case
VAR
    con : FB_EipConnect;
    dis : FB_EipDisconnect;
    sta : FB_EipStatus;
    lid : FB_EipListIdentity;
    ga  : FB_EipGetAttribute;
    sa  : FB_EipSetAttribute;
    st : INT;
    waitN : INT;
    mask AT %QD0 : UDINT;
    hdl : UDINT;
END_VAR
    IF st = 0 THEN
        mask := 0;
        con.Execute := TRUE;
        con.RemoteHost := '127.0.0.1';
        con.RemotePort := 14481;
        st := 1;
    END_IF;

    IF st = 1 THEN
        IF con.Done THEN
            hdl := con.SessionHdl;
            con.Execute := FALSE;
            mask := mask + 1;         // bit0: registered
            st := 2;
        END_IF;
        IF con.Error THEN mask := 16#DEAD; st := 99; END_IF;
    END_IF;

    IF st = 2 THEN
        waitN := waitN + 1;
        IF waitN >= 4 THEN
            sta.Execute := TRUE;
            sta.SessionHdl := hdl;
            st := 3;
        END_IF;
    END_IF;

    IF st = 3 THEN
        IF sta.Done THEN
            IF sta.SessionState = 1 AND sta.SessionId <> 0 THEN
                mask := mask + 2;             // bit1: session open
                sta.Execute := FALSE;
                lid.Execute := TRUE;
                lid.RemoteHost := '127.0.0.1';
                lid.RemotePort := 14481;
                st := 4;
            END_IF;
        END_IF;
        IF sta.Error THEN mask := 16#DEAD; st := 99; END_IF;
    END_IF;

    IF st = 4 THEN
        IF lid.Done THEN
            mask := mask + 4;                 // bit2: identity read
            lid.Execute := FALSE;
            ga.Execute := TRUE;
            ga.SessionHdl := hdl;
            ga.ClassId := 4;
            ga.InstanceId := 100;
            ga.AttributeId := 3;
            st := 5;
        END_IF;
        IF lid.Error THEN mask := 16#DEAD; st := 99; END_IF;
    END_IF;

    IF st = 5 THEN
        IF ga.Done THEN
            IF ga.ValueLen = 4 THEN
                mask := mask + 8;             // bit3: attr read (4B)
            END_IF;
            ga.Execute := FALSE;
            sa.Execute := TRUE;
            sa.SessionHdl := hdl;
            sa.ClassId := 4;
            sa.InstanceId := 100;
            sa.AttributeId := 3;
            sa.Value := 'ABCD';
            st := 6;
        END_IF;
        IF ga.Error THEN mask := 16#DEAD; st := 99; END_IF;
    END_IF;

    IF st = 6 THEN
        IF sa.Done THEN
            mask := mask + 16;                // bit4: attr written
            sa.Execute := FALSE;
            ga.Execute := TRUE;
            st := 7;
        END_IF;
        IF sa.Error THEN mask := 16#DEAD; st := 99; END_IF;
    END_IF;

    IF st = 7 THEN
        IF ga.Done THEN
            IF ga.Value = 'ABCD' THEN
                mask := mask + 32;            // bit5: readback ABCD
            END_IF;
            ga.Execute := FALSE;
            dis.Execute := TRUE;
            dis.SessionHdl := hdl;
            st := 8;
        END_IF;
        IF ga.Error THEN mask := 16#DEAD; st := 99; END_IF;
    END_IF;

    IF st = 8 THEN
        IF dis.Done THEN
            mask := mask + 64;                // bit6: disconnected
            st := 9;
        END_IF;
        IF dis.Error THEN mask := 16#DEAD; st := 99; END_IF;
    END_IF;

    con(); dis(); sta(); lid(); ga(); sa();
END_PROGRAM

(* ---- tc2_enocean_case.st ---- *)
// tc2_enocean_case.st — wired EnOcean ESP3 e2e over a PTY
// transceiver fake.  Open port, send a RADIO telegram (fake
// ACKs with RESPONSE + emits an inbound PTM radio), poll the
// receive, decode the PTM action, close.
PROGRAM tc2_enocean_case
VAR
    opn : FB_EnOceanOpen;
    cls : FB_EnOceanClose;
    snd : FB_EnOceanSendRadio;
    rx  : FB_EnOceanReceive;
    ptm : FB_EnOceanPtm100;
    st : INT;
    waitN : INT;
    mask AT %QD0 : UDINT;
    m2 : UDINT;
    diag AT %QD4 : UDINT;
    hdl : UDINT;
END_VAR
    diag := st;
    mask := m2;
    IF st = 0 THEN
        m2 := 0;
        opn.Execute := TRUE;
        opn.Path := '/tmp/eno_pty';
        st := 1;

    ELSIF st = 1 THEN
        IF opn.Done THEN
            hdl := opn.PortHdl;
            opn.Execute := FALSE;
            m2 := m2 OR 1;        // bit0: serial open
            snd.Execute := TRUE;
            snd.PortHdl := hdl;
            snd.Org := 16#F6;         // RPS
            snd.SenderId := 16#AABBCCDD;
            snd.DestId := 16#FFFFFFFF;
            snd.Data := 'x';
            st := 2;
        END_IF;
        IF opn.Error THEN diag := 1; m2 := 16#DE00 + 1; st := 99; END_IF;

    ELSIF st = 2 THEN
        IF snd.Done THEN
            m2 := m2 OR 2;        // bit1: radio frame sent
            snd.Execute := FALSE;
            rx.Execute := TRUE;
            rx.PortHdl := hdl;
            st := 3;
        END_IF;
        IF snd.Error THEN diag := 2; m2 := 16#DE00 + 2; st := 99; END_IF;

    // poll for the inbound radio telegram (fake emits after it
    // sees our transmit; RESPONSE packet may arrive first and
    // must be skipped, PTYPE=2)
    ELSIF st = 3 THEN
        waitN := waitN + 1;
        IF rx.Telegram THEN
            IF rx.PacketType = 1 AND rx.Org = 16#F6 AND rx.SenderId = 16#00112233 THEN
                m2 := m2 OR 4;    // bit2: radio decoded
                ptm.Execute := TRUE;
                ptm.Org := rx.Org;
                ptm.B0 := rx.Data0;
                st := 4;
            END_IF;
        END_IF;
        IF rx.Error THEN diag := 3; m2 := 16#DE00 + 3; st := 99; END_IF;
        IF waitN > 80 THEN diag := 4; m2 := 16#DE00 + 4; st := 99; END_IF;

    ELSIF st = 4 THEN
        rx.Execute := FALSE;
        IF ptm.Done AND ptm.IsPtm AND ptm.Pressed AND ptm.Act = 2 THEN
            m2 := m2 OR 8;        // bit3: PTM decode
            cls.Execute := TRUE;
            cls.PortHdl := hdl;
            st := 5;
        END_IF;

    ELSIF st = 5 THEN
        IF cls.Done THEN
            m2 := m2 OR 16;       // bit4: close ok
            st := 6;
        END_IF;
        IF cls.Error THEN diag := 5; m2 := 16#DE00 + 5; st := 99; END_IF;
    END_IF;

    opn(); cls(); snd(); rx(); ptm();
END_PROGRAM

(* ---- tc2_filter_case.st ---- *)
// tc2_filter_case.st — Tc2_Filter surface e2e: PT1 step response,
// PID tracking, limit clamp, average, ramp — pure-ST blocks.
PROGRAM tc2_filter_case
VAR
    lim : FB_Limit;
    pt1 : FB_PT1;
    pid : FB_PID;
    avg : FB_Average;
    rmp : FB_Ramp;
    st : INT;
    n : INT;
    mask AT %QD0 : UDINT;
END_VAR
    IF st = 0 THEN
        mask := 0;
        n := 0;
        lim.Execute := TRUE;
        pt1.Execute := TRUE;
        pid.Execute := TRUE;
        avg.Execute := TRUE;
        rmp.Execute := TRUE;
        pt1.Input := 1.0;   pt1.Kp := 1.0;  pt1.Tn := 0.5;  pt1.CycleTime := 0.1;
        pid.Setpoint := 1.0; pid.Actual := 0.0;
        pid.Kp := 2.0; pid.Tn := 0.5; pid.Tv := 0.0;
        pid.OutMin := -10.0; pid.OutMax := 10.0; pid.CycleTime := 0.1;
        avg.Input := 2.0; avg.N := 4;
        rmp.Setpoint := 3.0; rmp.SlewRate := 2.0; rmp.CycleTime := 0.1;
        lim.Input := 5.0; lim.Low := 0.0; lim.High := 3.0;
        st := 1;
    END_IF;

    IF st = 1 THEN
        IF lim.Done THEN
            IF lim.Output = 3.0 THEN mask := mask + 1; END_IF; // clamped
            st := 2;
        END_IF;
    END_IF;
    IF st = 2 THEN
        IF pt1.Done THEN
            n := n + 1;
            IF n > 20 THEN
                IF pt1.Output > 0.8 THEN mask := mask + 2; END_IF; // settles ~1
                n := 0;
                st := 3;
            END_IF;
        END_IF;
    END_IF;
    IF st = 3 THEN
        IF pid.Done THEN
            n := n + 1;
            IF n > 20 THEN
                IF pid.Output > 0.0 THEN mask := mask + 4; END_IF; // drives +
                n := 0;
                st := 4;
            END_IF;
        END_IF;
    END_IF;
    IF st = 4 THEN
        IF avg.Done THEN
            n := n + 1;
            IF n > 6 THEN
                IF avg.Output > 1.9 THEN mask := mask + 8; END_IF; // ~2.0
                n := 0;
                st := 5;
            END_IF;
        END_IF;
    END_IF;
    IF st = 5 THEN
        IF rmp.Done THEN
            n := n + 1;
            IF n > 40 THEN
                IF rmp.Output > 2.0 THEN mask := mask + 16; END_IF; // ramps
                n := 0;
                st := 6;
            END_IF;
        END_IF;
    END_IF;

    lim(); pt1(); pid(); avg(); rmp();
END_PROGRAM

(* ---- tc2_genibus_case.st ---- *)
// tc2_genibus_case.st — wired GENIbus e2e over a PTY slave
// fake (unit 0x20).  Open, ping -> ack, GET -> APDU reply,
// close.
PROGRAM tc2_genibus_case
VAR
    opn : FB_GenibusOpen;
    cls : FB_GenibusClose;
    png : FB_GENIbusPing;
    get : FB_GENIbusGet;
    rx  : FB_GENIbusReceive;
    st : INT;
    waitN : INT;
    mask AT %QD0 : UDINT;
    diag AT %QD4 : UDINT;
    hdl : UDINT;
END_VAR
    diag := st;
    IF st = 0 THEN
        mask := 0;
        opn.Execute := TRUE;
        opn.Path := '/tmp/gen_pty';
        st := 1;
    ELSIF st = 1 THEN
        IF opn.Done THEN
            hdl := opn.PortHdl;
            opn.Execute := FALSE;
            mask := mask OR 1;        // bit0: serial open
            png.Execute := TRUE;
            png.PortHdl := hdl;
            png.DestAddr := 16#20;
            png.SrcAddr := 0;
            st := 2;
        END_IF;
        IF opn.Error THEN diag := 16#D0; st := 99; END_IF;
    ELSIF st = 2 THEN
        IF png.Done THEN
            mask := mask OR 2;        // bit1: ping sent
            png.Execute := FALSE;
            rx.Execute := TRUE;
            rx.PortHdl := hdl;
            st := 3;
        END_IF;
        IF png.Error THEN diag := 16#D1; st := 99; END_IF;
    ELSIF st = 3 THEN
        waitN := waitN + 1;
        IF rx.Telegram THEN
            IF rx.SrcAddr = 16#20 THEN
                mask := mask OR 4;    // bit2: slave ack
                rx.Execute := FALSE;
                get.Execute := TRUE;
                get.PortHdl := hdl;
                get.DestAddr := 16#20;
                get.Item := 16#42;
                st := 4;
            END_IF;
        END_IF;
        IF rx.Error THEN diag := 16#D2; st := 99; END_IF;
        IF waitN > 80 THEN diag := 16#D3; st := 99; END_IF;
    ELSIF st = 4 THEN
        waitN := 0;
        IF get.Done THEN
            mask := mask OR 8;        // bit3: GET sent
            get.Execute := FALSE;
            rx.Execute := TRUE;
            st := 5;
        END_IF;
        IF get.Error THEN diag := 16#D4; st := 99; END_IF;
    ELSIF st = 5 THEN
        waitN := waitN + 1;
        IF rx.Telegram THEN
            IF rx.SrcAddr = 16#20 AND rx.ApduLen > 0 THEN
                mask := mask OR 16;   // bit4: APDU reply
                rx.Execute := FALSE;
                cls.Execute := TRUE;
                cls.PortHdl := hdl;
                st := 6;
            END_IF;
        END_IF;
        IF rx.Error THEN diag := 16#D5; st := 99; END_IF;
        IF waitN > 80 THEN diag := 16#D6; st := 99; END_IF;
    ELSIF st = 6 THEN
        IF cls.Done THEN
            mask := mask OR 32;       // bit5: close ok
            st := 7;
        END_IF;
        IF cls.Error THEN diag := 16#D7; st := 99; END_IF;
    END_IF;

    opn(); cls(); png(); get(); rx();
END_PROGRAM

(* ---- tc2_hvac_case.st ---- *)
// tc2_hvac_case.st — pure-ST e2e for tc2_hvac.
PROGRAM tc2_hvac_case
VAR
    ain : FB_HVACAnalogInput;
    aout : FB_HVACAnalogOutput;
    tp2 : FB_HVAC2PointActuator;
    tp3 : FB_HVAC3PointActuator;
    pump : FB_HVACCirculationPump;
    mot : FB_HVACMotor3Speed;
    mux : FB_HVACMux8;
    red : FB_HVACRedundancyCtrl;
    c2p : FB_HVAC2PointCtrl;
    stp : FB_HVACI_CtrlStep;
    pid : FB_HVACPIDCtrl;
    hcv : FB_HVACHeatingCurve;
    dmp : FB_HVACOutsideTempDamped;
    alm : FB_HVACAlarm;
    abp : FB_HVACAntiBlockingPump;
    blk : FB_HVACBlink;
    bar : FB_BARSetpointRoom;
    dhy : FB_BARDelayedHysteresis;
    st : INT;
    waitN : INT;
    mask AT %QD0 : UDINT;
    diag AT %QD4 : UDINT;
END_VAR
    diag := st;
    IF st = 0 THEN
        mask := 0;
        // analog input: 8000 of 0..16000 -> 0..50 = 25
        ain.Raw := 8000.0; ain.RawMin := 0.0; ain.RawMax := 16000.0;
        ain.EngMin := 0.0; ain.EngMax := 50.0;
        st := 1;
    ELSIF st = 1 THEN
        IF ain.Value > 24.9 AND ain.Value < 25.1 THEN mask := mask OR 1; END_IF;
        // 2-point ctrl: heating, actual below SP-hyst -> on
        c2p.bEnable := TRUE;
        c2p.fActual := 18.0; c2p.fSetpoint := 21.0; c2p.fHysteresis := 1.0;
        st := 2;
    ELSIF st = 2 THEN
        IF c2p.bOut THEN mask := mask OR 2; END_IF;
        // step ctrl: error 6 of 8 range, 4 stages -> 3 stages
        stp.bEnable := TRUE;
        stp.fActual := 14.0; stp.fSetpoint := 20.0;
        stp.fStepRange := 8.0; stp.nStages := 4;
        st := 3;
    ELSIF st = 3 THEN
        IF stp.bStage1 AND stp.bStage2 AND stp.bStage3 AND NOT stp.bStage4 THEN
            mask := mask OR 4;
        END_IF;
        // PID: error positive -> output above min
        pid.bEnable := TRUE;
        pid.fActual := 18.0; pid.fSetpoint := 22.0;
        pid.fKp := 2.0; pid.fTi := 0.0; pid.fTd := 0.0;
        pid.fOutMin := 0.0; pid.fOutMax := 100.0;
        pid.CycleTime := 0.1;
        st := 4;
    ELSIF st = 4 THEN
        IF pid.fOut > 5.0 THEN mask := mask OR 8; END_IF;
        // heating curve: outside -10, design -15, room 20
        // flow = 30 + (80-30) * (20-(-10)) / (20-(-15)) = 30+50*30/35 ≈ 72.86
        hcv.bEnable := TRUE;
        hcv.fOutsideTemp := -10.0; hcv.fOutsideMin := -15.0;
        hcv.fRoomTemp := 20.0; hcv.fSpMin := 30.0; hcv.fSpMax := 80.0;
        st := 5;
    ELSIF st = 5 THEN
        IF hcv.fFlowSp > 70.0 AND hcv.fFlowSp < 76.0 THEN mask := mask OR 16; END_IF;
        // motor3 speed 2 -> out2 only
        mot.bEnable := TRUE; mot.Speed := 2;
        mux.Sel := 3; mux.In3 := 42.0;
        st := 6;
    ELSIF st = 6 THEN
        IF mot.bOut2 AND NOT mot.bOut1 AND NOT mot.bOut3 THEN mask := mask OR 32; END_IF;
        IF mux.Out = 42.0 THEN mask := mask OR 64; END_IF;
        // redundancy: need 2, fault1 -> out2+out3
        red.bEnable := TRUE; red.Required := 2;
        red.bFault1 := TRUE;
        st := 7;
    ELSIF st = 7 THEN
        IF red.bOut2 AND red.bOut3 AND NOT red.bOut1 THEN mask := mask OR 128; END_IF;
        // alarm: value over limit 1s delay
        alm.bEnable := TRUE;
        alm.fValue := 10.0; alm.fLimit := 5.0; alm.fHysteresis := 1.0;
        alm.tDelay := 0.5; alm.CycleTime := 0.1;
        waitN := 0;
        st := 8;
    ELSIF st = 8 THEN
        waitN := waitN + 1;
        IF alm.bAlarm THEN mask := mask OR 256; st := 9; END_IF;
        IF waitN > 40 THEN diag := 16#E8; st := 99; END_IF;
    ELSIF st = 9 THEN
        // anti-blocking: idle pump exercises after tIdle
        abp.bEnable := TRUE; abp.bDemand := FALSE;
        abp.tIdle := 0.5; abp.tRunTime := 0.4; abp.CycleTime := 0.1;
        waitN := 0;
        st := 10;
    ELSIF st = 10 THEN
        waitN := waitN + 1;
        IF abp.bExercise THEN mask := mask OR 512; st := 11; END_IF;
        IF waitN > 40 THEN diag := 16#E9; st := 99; END_IF;
    ELSIF st = 11 THEN
        // blinker toggles
        blk.bEnable := TRUE; blk.tOn := 0.2; blk.tOff := 0.2;
        blk.CycleTime := 0.1;
        waitN := 0;
        st := 12;
    ELSIF st = 12 THEN
        waitN := waitN + 1;
        IF blk.bOut THEN mask := mask OR 1024; st := 13; END_IF;
        IF waitN > 40 THEN diag := 16#EA; st := 99; END_IF;
    ELSIF st = 13 THEN
        // bar setpoint: base 21 + shift 5 clamped to +3
        bar.bEnable := TRUE;
        bar.fBaseSp := 21.0; bar.fShift := 5.0; bar.fShiftMax := 3.0;
        // delayed hysteresis
        dhy.bEnable := TRUE;
        dhy.fValue := 10.0; dhy.fOn := 5.0; dhy.fOff := 2.0;
        dhy.tOnDelay := 0.0; dhy.tOffDelay := 0.0;
        dhy.CycleTime := 0.1;
        st := 14;
    ELSIF st = 14 THEN
        IF bar.fSetpoint = 24.0 THEN mask := mask OR 2048; END_IF;
        waitN := waitN + 1;
        IF dhy.bOut THEN mask := mask OR 4096; st := 15; END_IF;
        IF waitN > 40 THEN diag := 16#EB; st := 99; END_IF;
    ELSIF st = 15 THEN
        // 3-point actuator drives open
        tp3.bEnable := TRUE; tp3.bOpen := TRUE;
        tp3.tRun := 1.0; tp3.CycleTime := 0.1;
        waitN := 0;
        st := 16;
    ELSIF st = 16 THEN
        waitN := waitN + 1;
        IF tp3.Position > 50.0 THEN mask := mask OR 8192; st := 17; END_IF;
        IF waitN > 60 THEN diag := 16#EC; st := 99; END_IF;
    ELSIF st = 17 THEN
        // circulation pump: lead1 faulted -> pump2 runs
        pump.bEnable := TRUE; pump.bDemand := TRUE;
        pump.bFault1 := TRUE;
        st := 18;
    ELSIF st = 18 THEN
        IF pump.bPump2 AND NOT pump.bPump1 THEN mask := mask OR 16384; END_IF;
        // 2-point actuator: open command, endswitch ok
        tp2.bEnable := TRUE; tp2.bIn := TRUE;
        tp2.bLimitSwitchOpen := FALSE; tp2.bLimitSwitchClose := TRUE;
        tp2.tRun := 1.0; tp2.CycleTime := 0.1;
        waitN := 0;
        st := 19;
    ELSIF st = 19 THEN
        waitN := waitN + 1;
        IF tp2.Position > 50.0 THEN mask := mask OR 32768; st := 20; END_IF;
        IF waitN > 60 THEN diag := 16#ED; st := 99; END_IF;
    END_IF;

    ain(); aout(); tp2(); tp3(); pump(); mot(); mux(); red();
    c2p(); stp(); pid(); hcv(); dmp(); alm(); abp(); blk();
    bar(); dhy();
END_PROGRAM

(* ---- tc2_iec61850_brcb_case.st ---- *)
// tc2_iec61850_brcb_case.st — IEC 61850 buffered-RCB e2e over the
// fake IED: GetRCBValues on the $BR$ URCB twin, SetRCBValues enable,
// dataset write, dchg InformationReport via report poll, PurgeBuf,
// disable, disconnect.
PROGRAM tc2_iec61850_brcb_case
VAR
    con : FB_Iec61850Connect;
    dis : FB_Iec61850Disconnect;
    rget : FB_Iec61850RCBGet;
    rset : FB_Iec61850RCBSet;
    poll : FB_Iec61850ReportPoll;
    wr  : FB_Iec61850Write;
    st : INT;
    waitN : INT;
    mask AT %QD0 : UDINT;
    hdl : UDINT;
    rcbref : STRING[127];
    rep : STRING[255];
END_VAR
    IF st = 0 THEN
        mask := 0;
        rcbref := 'tetherIEDtetherTestLD/LLN0$$BR$$bufrcb';
        con.Execute := TRUE;
        con.RemoteHost := '127.0.0.1';
        con.RemotePort := 11020;
        st := 1;
    ELSIF st = 1 THEN
        IF con.Done THEN
            hdl := con.ConnectionHdl;
            con.Execute := FALSE;
            mask := mask + 1;
            rget.Execute := TRUE;
            rget.ConnectionHdl := hdl;
            rget.RcbRef := rcbref;
            st := 2;
        END_IF;
        IF con.Error THEN mask := 16#DEAD; st := 99; END_IF;
    ELSIF st = 2 THEN
        IF rget.Done THEN
            rget.Execute := FALSE;
            // rptId 'rptBuf', confRev 1, buffered, dchg+gi trgOps
            IF LEN(rget.RptId) = 6 AND FIND(rget.RptId, 'rptBuf') = 1
               AND rget.ConfRev = 1 AND rget.Buffered
               AND (rget.TrgOps AND 16#11) <> 0 THEN
                mask := mask + 2;
                rset.Execute := TRUE;
                rset.ConnectionHdl := hdl;
                rset.RcbRef := rcbref;
                rset.Flags := 1;      // rptEna
                st := 3;
            ELSE
                mask := 16#DEAD; st := 99;
            END_IF;
        END_IF;
        IF rget.Error THEN mask := 16#DEAD; st := 99; END_IF;
    ELSIF st = 3 THEN
        IF rset.Done THEN
            rset.Execute := FALSE;
            mask := mask + 4;
            wr.Execute := TRUE;
            wr.ConnectionHdl := hdl;
            wr.Domain := 'tetherIEDtetherTestLD';
            wr.Item := 'LLN0.SetPt.setMag.f#SP';
            wr.Value := '3.5';
            st := 4;
        END_IF;
        IF rset.Error THEN mask := 16#DEAD; st := 99; END_IF;
    ELSIF st = 4 THEN
        IF wr.Done THEN
            wr.Execute := FALSE;
            mask := mask + 8;
            waitN := 0;
            st := 5;
        END_IF;
        IF wr.Error THEN mask := 16#DEAD; st := 99; END_IF;
    ELSIF st = 5 THEN
        poll.Execute := TRUE;
        poll.ConnectionHdl := hdl;
        st := 50;
    ELSIF st = 50 THEN
        IF poll.Done THEN
            poll.Execute := FALSE;
            rep := poll.Report;
            // dchg report: dataset name + changed value only; older
            // buffered reports may still be queued, keep polling
            // until the post-write report shows up.
            IF poll.ReportBytes > 0
               AND FIND(rep, 'measds') > 0 AND FIND(rep, '3.5') > 0 THEN
                mask := mask + 16;
                waitN := 0;
                st := 64;             // arm integrity-report poll
            ELSIF waitN > 80 THEN
                mask := 16#DEAD; st := 99;
            ELSE
                waitN := waitN + 1;
                st := 5;
            END_IF;
        END_IF;
        IF poll.Error THEN mask := 16#DEAD; st := 99; END_IF;
    ELSIF st = 64 THEN
        poll.Execute := TRUE;
        poll.ConnectionHdl := hdl;
        st := 63;
    ELSIF st = 63 THEN
        // reap the unsolicited integrity report (intgPd=200 ms)
        IF poll.Done THEN
            poll.Execute := FALSE;
            rep := poll.Report;
            // integrity report: dataset name + every element value
            IF poll.ReportBytes > 0
               AND FIND(rep, 'measds') > 0 AND FIND(rep, '42') > 0
               AND FIND(rep, '3.5') > 0 THEN
                mask := mask + 256;
                rset.Execute := TRUE;
                rset.ConnectionHdl := hdl;
                rset.RcbRef := rcbref;
                rset.Flags := 0;      // disable (PurgeBuf needs disabled)
                st := 60;
            ELSIF waitN > 120 THEN
                mask := 16#DEAD; st := 99;
            ELSE
                waitN := waitN + 1;
                st := 64;             // re-arm via arm state
            END_IF;
        END_IF;
        IF poll.Error THEN mask := 16#DEAD; st := 99; END_IF;
    ELSIF st = 60 THEN
        IF rset.Done THEN
            rset.Execute := FALSE;
            mask := mask + 32;
            st := 62;
        END_IF;
        IF rset.Error THEN mask := 16#DEAD; st := 99; END_IF;
    ELSIF st = 62 THEN
        // arm the disable write (Execute was low last scan)
        rset.Execute := TRUE;
        rset.ConnectionHdl := hdl;
        rset.RcbRef := rcbref;
        rset.Flags := 8;      // PurgeBuf while disabled
        st := 61;
    ELSIF st = 61 THEN
        IF rset.Done THEN
            rset.Execute := FALSE;
            mask := mask + 64;
            dis.Execute := TRUE;
            dis.ConnectionHdl := hdl;
            st := 7;
        END_IF;
        IF rset.Error THEN mask := 16#DEAD; st := 99; END_IF;
    ELSIF st = 7 THEN
        IF dis.Done THEN
            dis.Execute := FALSE;
            mask := mask + 128;
            st := 99;
        END_IF;
        IF dis.Error THEN mask := 16#DEAD; END_IF;
    ELSIF st = 99 THEN
        // terminal
    END_IF
    con(); dis(); rget(); rset(); wr(); poll();
END_PROGRAM

(* ---- tc2_iec61850_case.st ---- *)
// tc2_iec61850_case.st — IEC 61850 client e2e over the fake IED.
// Connect+associate, read, write, GetNameList, disconnect.
PROGRAM tc2_iec61850_case
VAR
    con : FB_Iec61850Connect;
    dis : FB_Iec61850Disconnect;
    sta : FB_Iec61850Status;
    rd  : FB_Iec61850Read;
    wr  : FB_Iec61850Write;
    gnl : FB_Iec61850GetNameList;
    st : INT;
    waitN : INT;
    mask AT %QD0 : UDINT;
    hdl : UDINT;
END_VAR
    IF st = 0 THEN
        mask := 0;
        con.Execute := TRUE;
        con.RemoteHost := '127.0.0.1';
        con.RemotePort := 11020;
        st := 1;
    END_IF;

    IF st = 1 THEN
        IF con.Done THEN
            hdl := con.ConnectionHdl;
            con.Execute := FALSE;
            mask := mask + 1;         // bit0: associated
            st := 2;
        END_IF;
        IF con.Error THEN mask := 16#DEAD; st := 99; END_IF;
    END_IF;

    IF st = 2 THEN
        waitN := waitN + 1;
        IF waitN >= 4 THEN
            sta.Execute := TRUE;
            sta.ConnectionHdl := hdl;
            st := 3;
        END_IF;
    END_IF;

    IF st = 3 THEN
        IF sta.Done THEN
            IF sta.ConnectionState = 1 THEN
                mask := mask + 2;             // bit1: association open
                sta.Execute := FALSE;
                rd.Execute := TRUE;
                rd.ConnectionHdl := hdl;
                rd.Domain := 'tetherIEDtetherTestLD';
                rd.Item := 'LLN0.Name.val';
                st := 4;
            END_IF;
        END_IF;
        IF sta.Error THEN mask := 16#DEAD; st := 99; END_IF;
    END_IF;

    IF st = 4 THEN
        IF rd.Done THEN
            mask := mask + 4;                 // bit2: read issued
            rd.Execute := FALSE;
            rd.ConnectionHdl := hdl;
            rd.Domain := 'tetherIEDtetherTestLD';
            rd.Item := 'LLN0.Health.stVal';
            st := 5;
        END_IF;
        IF rd.Error THEN mask := 16#DEAD; st := 99; END_IF;
    END_IF;

    IF st = 5 THEN
        IF rd.Done THEN
            mask := mask + 8;                 // bit3: read stVal
            rd.Execute := FALSE;
            wr.Execute := TRUE;
            wr.ConnectionHdl := hdl;
            wr.Domain := 'tetherIEDtetherTestLD';
            wr.Item := 'LLN0.Health.stVal';
            wr.Value := '9';
            st := 6;
        END_IF;
        IF rd.Error THEN mask := 16#DEAD; st := 99; END_IF;
    END_IF;

    IF st = 6 THEN
        // write to a read-only stVal must report an MMS access error —
        // that verifies the write path returns a real server error
        IF wr.Error THEN
            mask := mask + 16;                // bit4: write path errors
            wr.Execute := FALSE;
            gnl.Execute := TRUE;
            gnl.ConnectionHdl := hdl;
            gnl.Domain := 'tetherIEDtetherTestLD';
            st := 7;
        END_IF;
        IF wr.Done THEN mask := 16#DEAD; st := 99; END_IF;
    END_IF;

    IF st = 7 THEN
        IF gnl.Done THEN
            mask := mask + 32;                // bit5: namelist
            gnl.Execute := FALSE;
            dis.Execute := TRUE;
            dis.ConnectionHdl := hdl;
            st := 8;
        END_IF;
        IF gnl.Error THEN mask := 16#DEAD; st := 99; END_IF;
    END_IF;

    IF st = 8 THEN
        IF dis.Done THEN
            mask := mask + 64;                // bit6: released
            st := 9;
        END_IF;
        IF dis.Error THEN mask := 16#DEAD; st := 99; END_IF;
    END_IF;

    con(); dis(); sta(); rd(); wr(); gnl();
END_PROGRAM

(* ---- tc2_iec61850_ctl_case.st ---- *)
// tc2_iec61850_ctl_case.st — IEC 61850 controllable-object e2e over
// the fake IED's SWI1 BSC (SBO normal + cancel): bare operate is
// rejected, select -> operate(true) -> stVal verifies, select ->
// cancel -> stVal unchanged, disconnect.
PROGRAM tc2_iec61850_ctl_case
VAR
    con : FB_Iec61850Connect;
    dis : FB_Iec61850Disconnect;
    ctl : FB_Iec61850Control;
    cpol : FB_Iec61850ControlPoll;
    rd  : FB_Iec61850Read;
    st : INT;
    waitN : INT;
    mask AT %QD0 : UDINT;
    hdl : UDINT;
    cref : STRING[127];
    sval : STRING[255];
END_VAR
    IF st = 0 THEN
        mask := 0;
        cref := 'tetherIEDtetherTestLD/LLN0.SWI1';
        con.Execute := TRUE;
        con.RemoteHost := '127.0.0.1';
        con.RemotePort := 11020;
        st := 1;
    ELSIF st = 1 THEN
        IF con.Done THEN
            hdl := con.ConnectionHdl;
            con.Execute := FALSE;
            mask := mask + 1;
            // bare operate without select must be rejected by the
            // SBO server (async CommandTermination- expected)
            ctl.Execute := TRUE;
            ctl.ConnectionHdl := hdl;
            ctl.ObjectRef := cref;
            ctl.Mode := 3;              // operate
            ctl.CtlValue := 'true';
            st := 20;
        END_IF;
        IF con.Error THEN mask := 16#DEAD; st := 99; END_IF;
    ELSIF st = 20 THEN
        IF ctl.Done THEN
            ctl.Execute := FALSE;
            mask := mask + 2;           // command accepted for tx
            waitN := 0;
            st := 21;
        END_IF;
        IF ctl.Error THEN mask := 16#DEAD; st := 99; END_IF;
    ELSIF st = 21 THEN
        cpol.Execute := TRUE;
        cpol.ConnectionHdl := hdl;
        st := 22;
    ELSIF st = 22 THEN
        IF cpol.Done THEN
            cpol.Execute := FALSE;
            // expect a pending operate termination with success=0
            IF cpol.Pending AND NOT cpol.Success
               AND cpol.EvType = 1 THEN
                mask := mask + 4;
                ctl.Execute := TRUE;
                ctl.ConnectionHdl := hdl;
                ctl.ObjectRef := cref;
                ctl.Mode := 1;          // select
                ctl.CtlValue := '';
                st := 23;
            ELSIF waitN > 100 THEN
                mask := 16#DEAD; st := 99;
            ELSE
                waitN := waitN + 1;
                st := 21;
            END_IF;
        END_IF;
        IF cpol.Error THEN mask := 16#DEAD; st := 99; END_IF;
    ELSIF st = 23 THEN
        IF ctl.Done THEN
            ctl.Execute := FALSE;
            mask := mask + 8;
            waitN := 0;
            st := 24;
        END_IF;
        IF ctl.Error THEN mask := 16#DEAD; st := 99; END_IF;
    ELSIF st = 24 THEN
        cpol.Execute := TRUE;
        cpol.ConnectionHdl := hdl;
        st := 25;
    ELSIF st = 25 THEN
        IF cpol.Done THEN
            cpol.Execute := FALSE;
            // select termination: type 0, success
            IF cpol.Pending AND cpol.Success AND cpol.EvType = 0 THEN
                mask := mask + 16;
                ctl.Execute := TRUE;
                ctl.ConnectionHdl := hdl;
                ctl.ObjectRef := cref;
                ctl.Mode := 3;          // operate
                ctl.CtlValue := 'true';
                st := 26;
            ELSIF waitN > 100 THEN
                mask := 16#DEAD; st := 99;
            ELSE
                waitN := waitN + 1;
                st := 24;
            END_IF;
        END_IF;
        IF cpol.Error THEN mask := 16#DEAD; st := 99; END_IF;
    ELSIF st = 26 THEN
        IF ctl.Done THEN
            ctl.Execute := FALSE;
            mask := mask + 32;
            waitN := 0;
            st := 27;
        END_IF;
        IF ctl.Error THEN mask := 16#DEAD; st := 99; END_IF;
    ELSIF st = 27 THEN
        cpol.Execute := TRUE;
        cpol.ConnectionHdl := hdl;
        st := 28;
    ELSIF st = 28 THEN
        IF cpol.Done THEN
            cpol.Execute := FALSE;
            // operate termination: type 1, success
            IF cpol.Pending AND cpol.Success AND cpol.EvType = 1 THEN
                mask := mask + 64;
                rd.Execute := TRUE;
                rd.ConnectionHdl := hdl;
                rd.Domain := 'tetherIEDtetherTestLD';
                rd.Item := 'LLN0.SWI1.valWTr.posVal#ST';
                st := 29;
            ELSIF waitN > 100 THEN
                mask := 16#DEAD; st := 99;
            ELSE
                waitN := waitN + 1;
                st := 27;
            END_IF;
        END_IF;
        IF cpol.Error THEN mask := 16#DEAD; st := 99; END_IF;
    ELSIF st = 29 THEN
        IF rd.Done THEN
            rd.Execute := FALSE;
            sval := rd.Value;
            // boolean stVal reads back as "1"
            IF FIND(sval, '1') > 0 THEN
                mask := mask + 128;
                // select again, then cancel: stVal must stay true
                ctl.Execute := TRUE;
                ctl.ConnectionHdl := hdl;
                ctl.ObjectRef := cref;
                ctl.Mode := 1;          // select
                ctl.CtlValue := '';
                st := 30;
            ELSE
                mask := 16#DEAD; st := 99;
            END_IF;
        END_IF;
        IF rd.Error THEN mask := 16#DEAD; st := 99; END_IF;
    ELSIF st = 30 THEN
        IF ctl.Done THEN
            ctl.Execute := FALSE;
            mask := mask + 256;
            waitN := 0;
            st := 31;
        END_IF;
        IF ctl.Error THEN mask := 16#DEAD; st := 99; END_IF;
    ELSIF st = 31 THEN
        cpol.Execute := TRUE;
        cpol.ConnectionHdl := hdl;
        st := 32;
    ELSIF st = 32 THEN
        IF cpol.Done THEN
            cpol.Execute := FALSE;
            IF cpol.Pending AND cpol.Success AND cpol.EvType = 0 THEN
                ctl.Execute := TRUE;
                ctl.ConnectionHdl := hdl;
                ctl.ObjectRef := cref;
                ctl.Mode := 4;          // cancel
                ctl.CtlValue := '';
                st := 33;
            ELSIF waitN > 100 THEN
                mask := 16#DEAD; st := 99;
            ELSE
                waitN := waitN + 1;
                st := 31;
            END_IF;
        END_IF;
        IF cpol.Error THEN mask := 16#DEAD; st := 99; END_IF;
    ELSIF st = 33 THEN
        IF ctl.Done THEN
            ctl.Execute := FALSE;
            mask := mask + 512;
            waitN := 0;
            st := 34;
        END_IF;
        IF ctl.Error THEN mask := 16#DEAD; st := 99; END_IF;
    ELSIF st = 34 THEN
        cpol.Execute := TRUE;
        cpol.ConnectionHdl := hdl;
        st := 35;
    ELSIF st = 35 THEN
        IF cpol.Done THEN
            cpol.Execute := FALSE;
            // cancel termination: type 2, success
            IF cpol.Pending AND cpol.Success AND cpol.EvType = 2 THEN
                mask := mask + 1024;
                rd.Execute := TRUE;
                rd.ConnectionHdl := hdl;
                rd.Domain := 'tetherIEDtetherTestLD';
                rd.Item := 'LLN0.SWI1.valWTr.posVal#ST';
                st := 36;
            ELSIF waitN > 100 THEN
                mask := 16#DEAD; st := 99;
            ELSE
                waitN := waitN + 1;
                st := 34;
            END_IF;
        END_IF;
        IF cpol.Error THEN mask := 16#DEAD; st := 99; END_IF;
    ELSIF st = 36 THEN
        IF rd.Done THEN
            rd.Execute := FALSE;
            sval := rd.Value;
            // cancel leaves stVal at the operated value (true)
            IF FIND(sval, '1') > 0 THEN
                mask := mask + 2048;
                // APC1: select -> operate(3.5) -> mxVal.f reads
                // back 3.5 through the structured ctlVal path
                cref := 'tetherIEDtetherTestLD/LLN0.APC1';
                ctl.Execute := TRUE;
                ctl.ConnectionHdl := hdl;
                ctl.ObjectRef := cref;
                ctl.Mode := 1;          // select
                ctl.CtlValue := '';
                st := 40;
            ELSE
                mask := 16#DEAD; st := 99;
            END_IF;
        END_IF;
        IF rd.Error THEN mask := 16#DEAD; st := 99; END_IF;
    ELSIF st = 40 THEN
        IF ctl.Done THEN
            ctl.Execute := FALSE;
            mask := mask + 4096;
            waitN := 0;
            st := 41;
        END_IF;
        IF ctl.Error THEN mask := 16#DEAD; st := 99; END_IF;
    ELSIF st = 41 THEN
        cpol.Execute := TRUE;
        cpol.ConnectionHdl := hdl;
        st := 42;
    ELSIF st = 42 THEN
        IF cpol.Done THEN
            cpol.Execute := FALSE;
            IF cpol.Pending AND cpol.Success AND cpol.EvType = 0 THEN
                ctl.Execute := TRUE;
                ctl.ConnectionHdl := hdl;
                ctl.ObjectRef := cref;
                ctl.Mode := 3;          // operate
                ctl.CtlValue := '3.5';
                st := 43;
            ELSIF waitN > 100 THEN
                mask := 16#DEAD; st := 99;
            ELSE
                waitN := waitN + 1;
                st := 41;
            END_IF;
        END_IF;
        IF cpol.Error THEN mask := 16#DEAD; st := 99; END_IF;
    ELSIF st = 43 THEN
        IF ctl.Done THEN
            ctl.Execute := FALSE;
            mask := mask + 8192;
            waitN := 0;
            st := 44;
        END_IF;
        IF ctl.Error THEN mask := 16#DEAD; st := 99; END_IF;
    ELSIF st = 44 THEN
        cpol.Execute := TRUE;
        cpol.ConnectionHdl := hdl;
        st := 45;
    ELSIF st = 45 THEN
        IF cpol.Done THEN
            cpol.Execute := FALSE;
            IF cpol.Pending AND cpol.Success AND cpol.EvType = 1 THEN
                rd.Execute := TRUE;
                rd.ConnectionHdl := hdl;
                rd.Domain := 'tetherIEDtetherTestLD';
                rd.Item := 'LLN0.APC1.mxVal.f#MX';
                st := 46;
            ELSIF waitN > 100 THEN
                mask := 16#DEAD; st := 99;
            ELSE
                waitN := waitN + 1;
                st := 44;
            END_IF;
        END_IF;
        IF cpol.Error THEN mask := 16#DEAD; st := 99; END_IF;
    ELSIF st = 46 THEN
        IF rd.Done THEN
            rd.Execute := FALSE;
            sval := rd.Value;
            IF sval = '3.5' THEN
                mask := mask + 16384;
                dis.Execute := TRUE;
                dis.ConnectionHdl := hdl;
                st := 7;
            ELSE
                mask := 16#DEAD; st := 99;
            END_IF;
        END_IF;
        IF rd.Error THEN mask := 16#DEAD; st := 99; END_IF;
    ELSIF st = 7 THEN
        IF dis.Done THEN
            dis.Execute := FALSE;
            mask := mask + 32768;
            st := 99;
        END_IF;
        IF dis.Error THEN mask := 16#DEAD; END_IF;
    ELSIF st = 99 THEN
        // terminal
    END_IF
    con(); dis(); ctl(); cpol(); rd();
END_PROGRAM

(* ---- tc2_iec61850_ds_case.st ---- *)
// tc2_iec61850_ds_case.st — IEC 61850 data-set e2e over the fake
// IED: GetDataSetDirectory + ReadDataSet on measds
// (Meas.instMag.f=42.5 MX + SetPt.setMag.f=1.0 SP), then
// WriteDataSet on writeds (SetPt.setMag.f + SetPt2.setMag.f, both SP)
// with a read-back verify, CreateDataSet/DeleteDataSet on the
// association-specific @dyn1 set, disconnect.
PROGRAM tc2_iec61850_ds_case
VAR
    con : FB_Iec61850Connect;
    dis : FB_Iec61850Disconnect;
    dsdir : FB_Iec61850DataSetDirectory;
    dsrd : FB_Iec61850DataSetRead;
    dswr : FB_Iec61850DataSetWrite;
    dscr : FB_Iec61850DataSetCreate;
    dsdell : FB_Iec61850DataSetDelete;
    st : INT;
    mask AT %QD0 : UDINT;
    hdl : UDINT;
    dsref : STRING[127];
    wdref : STRING[127];
    cref : STRING[127];
END_VAR
    IF st = 0 THEN
        mask := 0;
        dsref := 'tetherIEDtetherTestLD/LLN0.measds';
        wdref := 'tetherIEDtetherTestLD/LLN0.writeds';
        cref := '@dyn1';
        con.Execute := TRUE;
        con.RemoteHost := '127.0.0.1';
        con.RemotePort := 11020;
        st := 1;
    ELSIF st = 1 THEN
        IF con.Done THEN
            hdl := con.ConnectionHdl;
            con.Execute := FALSE;
            mask := mask + 1;
            dsdir.Execute := TRUE;
            dsdir.ConnectionHdl := hdl;
            dsdir.DataSetRef := dsref;
            st := 2;
        END_IF;
        IF con.Error THEN mask := 16#DEAD; st := 99; END_IF;
    ELSIF st = 2 THEN
        IF dsdir.Done THEN
            dsdir.Execute := FALSE;
            // two members: the MX instMag.f and SP setMag.f FCDAs
            IF dsdir.ElementCount = 2
               AND FIND(dsdir.Names, 'Meas') > 0
               AND FIND(dsdir.Names, 'SetPt') > 0 THEN
                mask := mask + 2;
            END_IF;
            dsrd.Execute := TRUE;
            dsrd.ConnectionHdl := hdl;
            dsrd.DataSetRef := dsref;
            st := 3;
        END_IF;
        IF dsdir.Error THEN mask := 16#DEAD; st := 99; END_IF;
    ELSIF st = 3 THEN
        IF dsrd.Done THEN
            dsrd.Execute := FALSE;
            // values: instMag.f=42.5, setMag.f=1.0
            IF dsrd.ElementCount = 2
               AND FIND(dsrd.Values, 'instMag') > 0
               AND FIND(dsrd.Values, '42.5') > 0
               AND FIND(dsrd.Values, 'setMag') > 0 THEN
                mask := mask + 4;
            END_IF;
            // WriteDataSet on the writable twin: stVal=9, setMag=7.25
            dswr.Execute := TRUE;
            dswr.ConnectionHdl := hdl;
            dswr.DataSetRef := wdref;
            dswr.Values := '9
7.25';
            st := 5;
        END_IF;
        IF dsrd.Error THEN mask := 16#DEAD; st := 99; END_IF;
    ELSIF st = 5 THEN
        IF dswr.Done THEN
            dswr.Execute := FALSE;
            mask := mask + 16;
            // read back the written dataset
            dsrd.Execute := TRUE;
            dsrd.ConnectionHdl := hdl;
            dsrd.DataSetRef := wdref;
            st := 6;
        END_IF;
        IF dswr.Error THEN mask := 16#DEAD; st := 99; END_IF;
    ELSIF st = 6 THEN
        IF dsrd.Done THEN
            dsrd.Execute := FALSE;
            IF dsrd.ElementCount = 2
               AND FIND(dsrd.Values, '9') > 0
               AND FIND(dsrd.Values, '7.25') > 0 THEN
                mask := mask + 32;
            END_IF;
            // create the association-specific @dyn1 data set with the
            // two writable members
            dscr.Execute := TRUE;
            dscr.ConnectionHdl := hdl;
            dscr.DataSetRef := cref;
            dscr.Elements := 'tetherIEDtetherTestLD/LLN0.SetPt.setMag.f[SP]
tetherIEDtetherTestLD/LLN0.SetPt2.setMag.f[SP]';
            st := 8;
        END_IF;
        IF dsrd.Error THEN mask := 16#DEAD; st := 99; END_IF;
    ELSIF st = 8 THEN
        IF dscr.Done THEN
            dscr.Execute := FALSE;
            mask := mask + 128;
            dsdir.Execute := TRUE;
            dsdir.ConnectionHdl := hdl;
            dsdir.DataSetRef := cref;
            st := 9;
        END_IF;
        IF dscr.Error THEN mask := 16#DEAD; st := 99; END_IF;
    ELSIF st = 9 THEN
        IF dsdir.Done THEN
            dsdir.Execute := FALSE;
            IF dsdir.ElementCount = 2 THEN
                mask := mask + 256;
            END_IF;
            dsdell.Execute := TRUE;
            dsdell.ConnectionHdl := hdl;
            dsdell.DataSetRef := cref;
            st := 10;
        END_IF;
        IF dsdir.Error THEN mask := 16#DEAD; st := 99; END_IF;
    ELSIF st = 10 THEN
        IF dsdell.Done THEN
            dsdell.Execute := FALSE;
            mask := mask + 512;
            // the deleted set must now be gone: directory errors
            dsdir.Execute := TRUE;
            dsdir.ConnectionHdl := hdl;
            dsdir.DataSetRef := cref;
            st := 11;
        END_IF;
        IF dsdell.Error THEN mask := 16#DEAD; st := 99; END_IF;
    ELSIF st = 11 THEN
        IF dsdir.Done THEN
            // unexpected success: the set survived deletion
            mask := 16#DEAD; st := 99;
        END_IF;
        IF dsdir.Error THEN
            dsdir.Execute := FALSE;
            mask := mask + 1024;
            dis.Execute := TRUE;
            dis.ConnectionHdl := hdl;
            st := 12;
        END_IF;
    ELSIF st = 12 THEN
        IF dis.Done THEN
            dis.Execute := FALSE;
            mask := mask + 2048;
            st := 99;
        END_IF;
        IF dis.Error THEN mask := 16#DEAD; st := 99; END_IF;
    END_IF;

    con(); dis(); dsdir(); dsrd(); dswr(); dscr(); dsdell();
END_PROGRAM

(* ---- tc2_iec61850_rcb_case.st ---- *)
// tc2_iec61850_rcb_case.st — IEC 61850 RCB e2e over the fake IED:
// GetRCBValues on the URCB, SetRCBValues enable, write a dataset
// member, receive the dchg InformationReport via report poll, send
// GI for a full-dataset report, disable, disconnect.
// dchg reports carry only changed elements ("-" for the rest);
// GI reports carry every dataset element.
PROGRAM tc2_iec61850_rcb_case
VAR
    con : FB_Iec61850Connect;
    dis : FB_Iec61850Disconnect;
    rget : FB_Iec61850RCBGet;
    rset : FB_Iec61850RCBSet;
    poll : FB_Iec61850ReportPoll;
    wr  : FB_Iec61850Write;
    st : INT;
    waitN : INT;
    mask AT %QD0 : UDINT;
    hdl : UDINT;
    rcbref : STRING[127];
    rep : STRING[255];
END_VAR
    IF st = 0 THEN
        mask := 0;
        rcbref := 'tetherIEDtetherTestLD/LLN0$$RP$$measurcb';
        con.Execute := TRUE;
        con.RemoteHost := '127.0.0.1';
        con.RemotePort := 11020;
        st := 1;
    ELSIF st = 1 THEN
        IF con.Done THEN
            hdl := con.ConnectionHdl;
            con.Execute := FALSE;
            mask := mask + 1;
            rget.Execute := TRUE;
            rget.ConnectionHdl := hdl;
            rget.RcbRef := rcbref;
            st := 2;
        END_IF;
        IF con.Error THEN mask := 16#DEAD; st := 99; END_IF;
    ELSIF st = 2 THEN
        IF rget.Done THEN
            rget.Execute := FALSE;
            // rptId 'rptMeas', confRev 1, unbuffered, dchg+gi trgOps
            IF LEN(rget.RptId) = 7 AND FIND(rget.RptId, 'rptMeas') = 1
               AND rget.ConfRev = 1 AND NOT rget.Buffered
               AND (rget.TrgOps AND 16#11) <> 0 THEN
                mask := mask + 2;
                rset.Execute := TRUE;
                rset.ConnectionHdl := hdl;
                rset.RcbRef := rcbref;
                rset.Flags := 1;      // rptEna
                st := 3;
            ELSE
                mask := 16#DEAD; st := 99;
            END_IF;
        END_IF;
        IF rget.Error THEN mask := 16#DEAD; st := 99; END_IF;
    ELSIF st = 3 THEN
        IF rset.Done THEN
            rset.Execute := FALSE;
            mask := mask + 4;
            wr.Execute := TRUE;
            wr.ConnectionHdl := hdl;
            wr.Domain := 'tetherIEDtetherTestLD';
            wr.Item := 'LLN0.SetPt.setMag.f#SP';
            wr.Value := '2.5';
            st := 4;
        END_IF;
        IF rset.Error THEN mask := 16#DEAD; st := 99; END_IF;
    ELSIF st = 4 THEN
        IF wr.Done THEN
            wr.Execute := FALSE;
            mask := mask + 8;
            waitN := 0;
            st := 5;
        END_IF;
        IF wr.Error THEN mask := 16#DEAD; st := 99; END_IF;
    ELSIF st = 5 THEN
        // arm one report poll per visit
        poll.Execute := TRUE;
        poll.ConnectionHdl := hdl;
        st := 50;
    ELSIF st = 50 THEN
        IF poll.Done THEN
            poll.Execute := FALSE;
            rep := poll.Report;
            IF poll.ReportBytes > 0 THEN
                // dchg report: dataset name + changed value only
                IF FIND(rep, 'measds') > 0 AND FIND(rep, '2.5') > 0 THEN
                    mask := mask + 16;
                END_IF;
                rset.Execute := TRUE;
                rset.ConnectionHdl := hdl;
                rset.RcbRef := rcbref;
                rset.Flags := 5;      // rptEna + GI
                st := 60;
            ELSIF waitN > 80 THEN
                mask := 16#DEAD; st := 99;
            ELSE
                waitN := waitN + 1;
                st := 5;
            END_IF;
        END_IF;
        IF poll.Error THEN mask := 16#DEAD; st := 99; END_IF;
    ELSIF st = 60 THEN
        IF rset.Done THEN
            rset.Execute := FALSE;
            mask := mask + 32;
            waitN := 0;
            poll.Execute := TRUE;
            poll.ConnectionHdl := hdl;
            st := 61;
        END_IF;
        IF rset.Error THEN mask := 16#DEAD; st := 99; END_IF;
    ELSIF st = 61 THEN
        // reap the GI report poll
        IF poll.Done THEN
            poll.Execute := FALSE;
            rep := poll.Report;
            IF poll.ReportBytes > 0 THEN
                // GI report: dataset name + every element value
                IF FIND(rep, 'measds') > 0 AND FIND(rep, '42') > 0
                   AND FIND(rep, '2.5') > 0 THEN
                    mask := mask + 64;
                END_IF;
                rset.Execute := TRUE;
                rset.ConnectionHdl := hdl;
                rset.RcbRef := rcbref;
                rset.Flags := 0;      // disable
                st := 62;
            ELSIF waitN > 80 THEN
                mask := 16#DEAD; st := 99;
            ELSE
                waitN := waitN + 1;
                poll.Execute := TRUE;   // re-arm for next visit
                st := 61;
            END_IF;
        END_IF;
        IF poll.Error THEN mask := 16#DEAD; st := 99; END_IF;
    ELSIF st = 62 THEN
        IF rset.Done THEN
            rset.Execute := FALSE;
            mask := mask + 128;
            dis.Execute := TRUE;
            dis.ConnectionHdl := hdl;
            st := 7;
        END_IF;
        IF rset.Error THEN mask := 16#DEAD; st := 99; END_IF;
    ELSIF st = 7 THEN
        IF dis.Done THEN
            dis.Execute := FALSE;
            mask := mask + 256;
            st := 99;
        END_IF;
        IF dis.Error THEN mask := 16#DEAD; END_IF;
    ELSIF st = 99 THEN
        // terminal
    END_IF
    con(); dis(); rget(); rset(); wr(); poll();
END_PROGRAM

(* ---- tc2_iofunctions_case.st ---- *)
// tc2_iofunctions_case.st — e2e for tc2_iofunctions (IOF general).
// The program declares three AT-bound "boxes"; the IOF blocks
// enumerate them by count, name and address.
PROGRAM tc2_iofunctions_case
VAR
    nBox : IOF_GetBoxCount;
    nDev : IOF_GetDeviceCount;
    byName : IOF_GetBoxAddrByName;
    byAddr : IOF_GetBoxNameByAddr;
    devName : IOF_GetDeviceName;
    devReset : IOF_DeviceReset;
    netId : IOF_GetDeviceNetId;
    in1 AT %IX0.0 : BOOL;
    out1 AT %QW2 : WORD;
    mem1 AT %MD4 : DWORD;
    st : INT;
    mask AT %QD0 : UDINT;
    diag AT %QD4 : UDINT;
END_VAR
    diag := st;
    IF st = 0 THEN
        mask := 0;
        nBox.bExecute := TRUE;
        st := 1;
    ELSIF st = 1 THEN
        nBox.bExecute := FALSE;
        IF nBox.bDone AND nBox.nCount = 5 THEN mask := mask OR 1; END_IF;
        nDev.bExecute := TRUE;
        st := 2;
    ELSIF st = 2 THEN
        nDev.bExecute := FALSE;
        IF nDev.bDone AND nDev.nCount = 1 THEN mask := mask OR 2; END_IF;
        byName.sName := 'out1';
        st := 3;
    ELSIF st = 3 THEN
        byName.bExecute := TRUE;
        st := 4;
    ELSIF st = 4 THEN
        byName.bExecute := FALSE;
        IF byName.bDone AND byName.nRegion = 1 AND byName.nAddr = 2 THEN
            mask := mask OR 4;
        END_IF;
        byAddr.nRegion := 2; byAddr.nAddr := 4;
        st := 5;
    ELSIF st = 5 THEN
        byAddr.bExecute := TRUE;
        st := 6;
    ELSIF st = 6 THEN
        byAddr.bExecute := FALSE;
        IF byAddr.bDone AND FIND(byAddr.sName, 'mem1') = 1 THEN
            mask := mask OR 8;
        END_IF;
        devName.nDevId := 0;
        st := 7;
    ELSIF st = 7 THEN
        devName.bExecute := TRUE;
        st := 8;
    ELSIF st = 8 THEN
        devName.bExecute := FALSE;
        IF devName.bDone AND FIND(devName.sName, 'Local') = 1 THEN
            mask := mask OR 16;
        END_IF;
        devReset.nDevId := 0;
        st := 9;
    ELSIF st = 9 THEN
        devReset.bExecute := TRUE;
        st := 10;
    ELSIF st = 10 THEN
        devReset.bExecute := FALSE;
        IF devReset.bError AND devReset.nErrId = 16#8001 THEN
            mask := mask OR 32;
        END_IF;
        netId.nDevId := 0;
        st := 11;
    ELSIF st = 11 THEN
        netId.bExecute := TRUE;
        st := 12;
    ELSIF st = 12 THEN
        netId.bExecute := FALSE;
        IF netId.bDone AND FIND(netId.sNetId, '127.0.0.1') = 1 THEN
            mask := mask OR 64;
        END_IF;
        st := 13;
    END_IF;
    nBox(); nDev(); byName(); byAddr(); devName(); devReset(); netId();
END_PROGRAM

(* ---- tc2_mbus_case.st ---- *)
// tc2_mbus_case.st — wired M-Bus master e2e over a PTY slave fake.
// Open, SND_NKE -> E5, REQ_UD2 -> data frame, close.
PROGRAM tc2_mbus_case
VAR
    opn : FB_MbusOpen;
    cls : FB_MbusClose;
    nke : FB_MbusShort;
    req : FB_MbusShort;
    rx  : FB_MbusReceive;
    st : INT;
    waitN : INT;
    mask AT %QD0 : UDINT;
    diag AT %QD4 : UDINT;
    hdl : UDINT;
END_VAR
    diag := 0;
    IF st = 0 THEN
        mask := 0;
        opn.Execute := TRUE;
        opn.Path := '/tmp/mbus_pty';
        st := 1;
    END_IF;

    IF st = 1 THEN
        IF opn.Done THEN
            hdl := opn.PortHdl;
            opn.Execute := FALSE;
            mask := mask + 1;         // bit0: serial open
            nke.Execute := TRUE;
            nke.PortHdl := hdl;
            nke.Control := 16#40;     // SND_NKE
            nke.Address := 1;
            st := 2;
        END_IF;
        IF opn.Error THEN diag := 1; mask := 16#DE00 + 1; st := 99; END_IF;
    END_IF;

    IF st = 2 THEN
        IF nke.Done THEN
            mask := mask + 2;         // bit1: NKE sent
            nke.Execute := FALSE;
            rx.Execute := TRUE;
            rx.PortHdl := hdl;
            st := 3;
        END_IF;
        IF nke.Error THEN diag := 2; mask := 16#DE00 + 2; st := 99; END_IF;
    END_IF;

    // poll for the slave's E5 ack
    IF st = 3 THEN
        waitN := waitN + 1;
        IF rx.Message THEN
            IF rx.Kind = 16#E5 THEN
                mask := mask + 4;     // bit2: E5 ack
            END_IF;
            rx.Execute := FALSE;
            req.Execute := TRUE;
            req.PortHdl := hdl;
            req.Control := 16#5B;     // REQ_UD2
            req.Address := 1;
            st := 4;
        END_IF;
        IF rx.Error THEN diag := 3; mask := 16#DE00 + 3; st := 99; END_IF;
        IF waitN > 40 THEN
            rx.Execute := FALSE;
            req.Execute := TRUE;
            req.PortHdl := hdl;
            req.Control := 16#5B;
            req.Address := 1;
            st := 4;
        END_IF;
    END_IF;

    IF st = 4 THEN
        IF req.Done THEN
            mask := mask + 8;         // bit3: REQ_UD2 sent
            req.Execute := FALSE;
            rx.Execute := TRUE;
            rx.PortHdl := hdl;
            waitN := 0;
            st := 5;
        END_IF;
        IF req.Error THEN diag := 4; mask := 16#DE00 + 4; st := 99; END_IF;
    END_IF;

    // poll for the slave's 68.. data frame
    IF st = 5 THEN
        waitN := waitN + 1;
        IF rx.Message THEN
            IF rx.Kind = 16#68 THEN
                mask := mask + 16;    // bit4: data frame
            END_IF;
            rx.Execute := FALSE;
            cls.Execute := TRUE;
            cls.PortHdl := hdl;
            st := 6;
        END_IF;
        IF rx.Error THEN diag := 5; mask := 16#DE00 + 5; st := 99; END_IF;
        IF waitN > 40 THEN
            rx.Execute := FALSE;
            cls.Execute := TRUE;
            cls.PortHdl := hdl;
            st := 6;
        END_IF;
    END_IF;

    IF st = 6 THEN
        IF cls.Done THEN
            mask := mask + 32;        // bit5: closed
            st := 7;
        END_IF;
        IF cls.Error THEN diag := 6; mask := 16#DE00 + 6; st := 99; END_IF;
    END_IF;

    opn(); cls(); nke(); req(); rx();
END_PROGRAM
